      R_f[3,4] := -0.60042000;
      R_f[3,5] := 0.30684051;
      R_f[3,6] := 0.39524430;
      R_f[3,7] := 0.11368765;
      R_f[3,8] := -0.22525014;
      R_f[3,9] := 0.40331784;
      R_f[3,10] := -0.22694421;
      R_f[3,11] := 0.08383388;
      R_f[3,12] := -0.06074797;
      R_f[3,13] := -0.18165708;
      R_f[3,14] := -0.04610621;
      R_f[3,15] := -0.62458295;
      R_f[3,16] := 0.00826784;
      R_f[3,17] := 0.13735548;
      R_f[3,18] := 0.04492014;
      R_f[3,19] := -0.30372253;
      R_f[3,20] := -0.08298360;
      R_f[3,21] := 0.43319181;
      R_f[3,22] := 0.03173294;
      R_f[3,23] := 0.26679260;
      R_f[3,24] := 0.19107546;
      R_f[3,25] := -0.13225158;
      R_f[3,26] := 0.04235943;
      R_f[3,27] := 0.73829132;
      R_f[3,28] := 0.57859170;
      R_f[3,29] := -0.07161227;
      R_f[3,30] := -0.07272696;
      R_f[3,31] := -0.50867581;
      R_f[4,0] := -1.08717740;
      R_f[4,1] := -0.04287297;
      R_f[4,2] := -0.19841136;
      R_f[4,3] := 0.24848095;
      R_f[4,4] := -0.64561760;
      R_f[4,5] := -0.20718722;
      R_f[4,6] := -0.05597278;
      R_f[4,7] := -0.16602105;
      R_f[4,8] := -0.29476261;
      R_f[4,9] := 0.47976902;
      R_f[4,10] := -0.05075360;
      R_f[4,11] := 0.14082003;
      R_f[4,12] := 0.06980632;
      R_f[4,13] := 0.33018085;
      R_f[4,14] := 0.04662931;
      R_f[4,15] := -0.07799391;
      R_f[4,16] := 0.00706400;
      R_f[4,17] := 0.13971923;
      R_f[4,18] := 0.03753237;
      R_f[4,19] := -0.02597110;
      R_f[4,20] := -0.60197109;
      R_f[4,21] := 0.04454581;
      R_f[4,22] := -0.13320792;
      R_f[4,23] := 0.31133512;
      R_f[4,24] := -0.16363572;
      R_f[4,25] := 0.41873544;
      R_f[4,26] := -0.52481866;
      R_f[4,27] := 0.06860130;
      R_f[4,28] := 0.00750138;
      R_f[4,29] := 0.00922540;
      R_f[4,30] := 0.12660387;
      R_f[4,31] := 0.11132577;
      R_f[5,0] := -0.08935551;
      R_f[5,1] := 0.00341007;
      R_f[5,2] := -0.36269036;
      R_f[5,3] := -0.05915058;
      R_f[5,4] := 0.65549088;
      R_f[5,5] := -0.45446295;
      R_f[5,6] := 0.02701634;
      R_f[5,7] := 0.33505848;
      R_f[5,8] := 0.33433130;
      R_f[5,9] := -0.11102643;
      R_f[5,10] := 0.04686662;
      R_f[5,11] := -0.11728232;
      R_f[5,12] := 0.09523005;
      R_f[5,13] := -0.37170398;
      R_f[5,14] := 0.00033050;
      R_f[5,15] := 0.02845602;
      R_f[5,16] := 0.42707691;
      R_f[5,17] := -0.06965928;
      R_f[5,18] := 0.01540217;
      R_f[5,19] := -0.15121390;
      R_f[5,20] := -0.04805366;
      R_f[5,21] := -0.18535455;
      R_f[5,22] := 0.32275927;
      R_f[5,23] := -0.19729009;
      R_f[5,24] := 0.34231305;
      R_f[5,25] := -0.36576355;
      R_f[5,26] := -0.06866702;
      R_f[5,27] := 0.00050627;
      R_f[5,28] := -0.22415085;
      R_f[5,29] := 0.21506223;
      R_f[5,30] := 0.28907591;
      R_f[5,31] := 0.08619282;
      R_f[6,0] := 0.18388480;
      R_f[6,1] := 0.05767936;
      R_f[6,2] := -0.22664715;
      R_f[6,3] := 0.10472890;
      R_f[6,4] := 0.13720502;
      R_f[6,5] := -0.05844464;
      R_f[6,6] := 0.40636781;
      R_f[6,7] := 0.23722953;
      R_f[6,8] := 0.06870923;
      R_f[6,9] := -0.07299573;
      R_f[6,10] := 0.39616698;
      R_f[6,11] := 0.05431297;
      R_f[6,12] := -0.15155350;
      R_f[6,13] := -0.13813569;
      R_f[6,14] := -0.10887969;
      R_f[6,15] := -0.06144879;
      R_f[6,16] := 0.08795995;
      R_f[6,17] := -0.14627954;
      R_f[6,18] := 0.07981436;
      R_f[6,19] := 0.18627544;
      R_f[6,20] := -0.07600380;
      R_f[6,21] := -0.34014723;
      R_f[6,22] := -0.54018772;
      R_f[6,23] := 0.29552394;
      R_f[6,24] := -0.10880617;
      R_f[6,25] := -0.08422133;
      R_f[6,26] := -0.24422757;
      R_f[6,27] := -0.03805847;
      R_f[6,28] := 0.16830419;
      R_f[6,29] := -0.18664716;
      R_f[6,30] := 0.20243780;
      R_f[6,31] := 0.07874886;
      R_f[7,0] := 0.28316271;
      R_f[7,1] := 0.13009299;
      R_f[7,2] := 0.04995405;
      R_f[7,3] := 0.14345303;
      R_f[7,4] := 0.08940059;
      R_f[7,5] := -0.04840774;
      R_f[7,6] := 0.17071612;
      R_f[7,7] := -0.00365471;
      R_f[7,8] := -0.10895292;
      R_f[7,9] := -0.20513341;
      R_f[7,10] := 0.09715845;
      R_f[7,11] := 0.05839429;
      R_f[7,12] := 0.04244281;
      R_f[7,13] := -0.05333439;
      R_f[7,14] := 0.10779919;
      R_f[7,15] := 0.00831443;
      R_f[7,16] := -0.02139841;
      R_f[7,17] := -0.27714881;
      R_f[7,18] := -0.13269936;
      R_f[7,19] := 0.38708043;
      R_f[7,20] := 0.02227914;
      R_f[7,21] := -0.12789786;
      R_f[7,22] := -0.21672793;
      R_f[7,23] := 0.04945551;
      R_f[7,24] := -0.12798266;
      R_f[7,25] := -0.08468608;
      R_f[7,26] := 0.04391497;
      R_f[7,27] := 0.04113905;
      R_f[7,28] := -0.10612858;
      R_f[7,29] := 0.10980094;
      R_f[7,30] := 0.06744546;
      R_f[7,31] := 0.15760666;
      R_f[8,0] := -0.09437604;
      R_f[8,1] := 0.10058102;
      R_f[8,2] := -0.39239755;
      R_f[8,3] := 0.07142383;
      R_f[8,4] := 0.32619441;
      R_f[8,5] := -0.29801306;
      R_f[8,6] := 0.17732149;
      R_f[8,7] := 0.39382425;
      R_f[8,8] := -0.25244871;
      R_f[8,9] := -0.78001058;
      R_f[8,10] := -0.09953760;
      R_f[8,11] := -0.01873088;
      R_f[8,12] := -0.12824003;
      R_f[8,13] := -0.04000987;
      R_f[8,14] := -0.32546988;
      R_f[8,15] := -0.07414734;
      R_f[8,16] := -0.15979169;
      R_f[8,17] := -0.16899861;
      R_f[8,18] := 0.11978716;
      R_f[8,19] := -0.29437670;
      R_f[8,20] := -0.07145600;
      R_f[8,21] := 0.37895897;
      R_f[8,22] := 0.60730362;
      R_f[8,23] := -0.01808002;
      R_f[8,24] := 0.18473065;
      R_f[8,25] := -0.63517946;
      R_f[8,26] := -0.07078326;
      R_f[8,27] := 0.01834848;
      R_f[8,28] := -0.27034160;
      R_f[8,29] := 0.03424344;
      R_f[8,30] := 0.17846985;
      R_f[8,31] := -0.10791938;
      R_f[9,0] := 0.50240064;
      R_f[9,1] := -0.19293827;
      R_f[9,2] := -0.14941828;
      R_f[9,3] := 0.30088151;
      R_f[9,4] := -0.22305536;
      R_f[9,5] := -0.20884813;
      R_f[9,6] := -0.52308059;
      R_f[9,7] := -0.08416846;
      R_f[9,8] := -0.31933308;
      R_f[9,9] := 0.74035096;
      R_f[9,10] := 0.06057476;
      R_f[9,11] := -0.31038794;
      R_f[9,12] := -0.02742688;
      R_f[9,13] := 0.24148650;
      R_f[9,14] := 0.22138420;
      R_f[9,15] := -0.50248486;
      R_f[9,16] := 0.03389943;
      R_f[9,17] := -0.15244213;
      R_f[9,18] := -0.23831080;
      R_f[9,19] := 0.18266003;
      R_f[9,20] := -0.04345531;
      R_f[9,21] := -0.16341494;
      R_f[9,22] := -0.13197300;
      R_f[9,23] := -0.01865776;
      R_f[9,24] := 0.46940479;
      R_f[9,25] := 0.06735769;
      R_f[9,26] := -0.33095923;
      R_f[9,27] := -0.07481478;
      R_f[9,28] := 0.30265671;
      R_f[9,29] := -0.02983976;
      R_f[9,30] := 0.11981419;
      R_f[9,31] := 0.43036476;
      R_f[10,0] := -0.16625722;
      R_f[10,1] := 0.18885586;
      R_f[10,2] := 0.30220106;
      R_f[10,3] := -0.08386957;
      R_f[10,4] := -0.50032878;
      R_f[10,5] := 0.08482117;
      R_f[10,6] := 0.13217595;
      R_f[10,7] := 0.13670275;
      R_f[10,8] := -0.27781987;
      R_f[10,9] := 0.05184001;
      R_f[10,10] := -0.32821399;
      R_f[10,11] := 0.06394526;
      R_f[10,12] := 0.70230156;
      R_f[10,13] := 0.14407636;
      R_f[10,14] := 0.21430548;
      R_f[10,15] := -0.13537307;
      R_f[10,16] := -0.70127255;
      R_f[10,17] := 0.08713871;
      R_f[10,18] := 0.49356794;
      R_f[10,19] := -0.33338264;
      R_f[10,20] := -0.14740926;
      R_f[10,21] := 0.22738504;
      R_f[10,22] := -0.12947781;
      R_f[10,23] := 0.15810163;
      R_f[10,24] := 0.01187740;
      R_f[10,25] := 0.16353421;
      R_f[10,26] := 0.49730638;
      R_f[10,27] := -0.06625025;
      R_f[10,28] := -0.15717453;
      R_f[10,29] := -0.17355147;
      R_f[10,30] := -0.03920694;
      R_f[10,31] := 0.30297169;
      R_f[11,0] := 0.12163632;
      R_f[11,1] := -0.16561009;
      R_f[11,2] := -0.63697898;
      R_f[11,3] := -0.12967597;
      R_f[11,4] := -0.15516940;
      R_f[11,5] := -0.43934959;
      R_f[11,6] := -0.84410143;
      R_f[11,7] := -0.15710612;
      R_f[11,8] := -0.91981030;
      R_f[11,9] := 0.10710724;
      R_f[11,10] := -0.25132748;
      R_f[11,11] := 0.77600086;
      R_f[11,12] := -0.20838273;
      R_f[11,13] := 0.32214221;
      R_f[11,14] := -0.02206153;
      R_f[11,15] := -0.39864928;
      R_f[11,16] := -0.17909747;
      R_f[11,17] := -0.08701507;
      R_f[11,18] := -0.16743112;
      R_f[11,19] := -0.54472065;
      R_f[11,20] := -0.58381855;
      R_f[11,21] := 0.13781570;
      R_f[11,22] := -0.65494400;
      R_f[11,23] := 0.08265506;
      R_f[11,24] := 0.11775696;
      R_f[11,25] := 0.86460680;
      R_f[11,26] := 0.22440501;
      R_f[11,27] := 0.10443961;
      R_f[11,28] := -0.11450481;
      R_f[11,29] := 0.10720722;
      R_f[11,30] := -0.14559385;
      R_f[11,31] := -0.41325647;
      R_f[12,0] := 0.08129373;
      R_f[12,1] := 0.20157976;
      R_f[12,2] := -0.09767752;
      R_f[12,3] := 0.11404920;
      R_f[12,4] := 0.06406736;
      R_f[12,5] := -0.10172413;
      R_f[12,6] := -0.62003994;
      R_f[12,7] := 0.29222506;
      R_f[12,8] := 0.09104837;
      R_f[12,9] := 0.02718525;
      R_f[12,10] := -0.17208911;
      R_f[12,11] := 0.11898477;
      R_f[12,12] := 0.14371057;
      R_f[12,13] := 0.07740860;
      R_f[12,14] := 0.03334129;
      R_f[12,15] := -0.34480530;
      R_f[12,16] := 0.11375867;
      R_f[12,17] := -0.16553403;
      R_f[12,18] := -0.03753847;
      R_f[12,19] := 0.42828915;
      R_f[12,20] := -0.23550081;
      R_f[12,21] := -0.64313370;
      R_f[12,22] := 0.11878636;
      R_f[12,23] := 0.06645127;
      R_f[12,24] := -0.05381826;
      R_f[12,25] := -0.06362370;
      R_f[12,26] := 0.14368635;
      R_f[12,27] := 0.03581888;
      R_f[12,28] := -0.27521226;
      R_f[12,29] := -0.06815766;
      R_f[12,30] := 0.05883517;
      R_f[12,31] := 0.01413656;
      R_f[13,0] := -0.09574396;
      R_f[13,1] := 0.30759236;
      R_f[13,2] := -0.40949357;
      R_f[13,3] := -0.30002195;
      R_f[13,4] := 0.62065625;
      R_f[13,5] := -0.06791952;
      R_f[13,6] := -0.10181803;
      R_f[13,7] := 0.06609505;
      R_f[13,8] := 0.45424458;
      R_f[13,9] := -0.32844600;
      R_f[13,10] := 0.17730820;
      R_f[13,11] := -0.15458618;
      R_f[13,12] := -0.16377521;
      R_f[13,13] := 0.12967198;
      R_f[13,14] := -0.18851388;
      R_f[13,15] := 0.08791368;
      R_f[13,16] := 0.19190530;
      R_f[13,17] := -0.03352485;
      R_f[13,18] := -0.24754001;
      R_f[13,19] := -0.03332811;
      R_f[13,20] := -0.22078300;
      R_f[13,21] := -0.27547061;
      R_f[13,22] := 0.77056712;
      R_f[13,23] := -0.11708862;
      R_f[13,24] := 0.38989946;
      R_f[13,25] := 0.12295369;
      R_f[13,26] := 0.01030140;
      R_f[13,27] := -0.10658067;
      R_f[13,28] := -0.25609714;
      R_f[13,29] := 0.09743972;
      R_f[13,30] := 0.57624507;
      R_f[13,31] := 0.09921760;
      R_f[14,0] := -0.46166307;
      R_f[14,1] := -0.38297445;
      R_f[14,2] := -0.34351581;
      R_f[14,3] := 0.50245303;
      R_f[14,4] := -0.47205976;
      R_f[14,5] := -0.04034173;
      R_f[14,6] := 0.19666021;
      R_f[14,7] := -0.15099366;
      R_f[14,8] := -0.23554653;
      R_f[14,9] := 0.44932032;
      R_f[14,10] := -0.24074826;
      R_f[14,11] := 0.29974288;
      R_f[14,12] := -0.44155741;
      R_f[14,13] := 0.83714885;
      R_f[14,14] := 0.18741892;
      R_f[14,15] := -0.21850257;
      R_f[14,16] := -0.12847616;
      R_f[14,17] := 0.06488960;
      R_f[14,18] := -0.00284800;
      R_f[14,19] := -0.31293416;
      R_f[14,20] := -0.07697109;
      R_f[14,21] := 0.38044301;
      R_f[14,22] := -0.48185810;
      R_f[14,23] := -0.07073558;
      R_f[14,24] := -0.99695712;
      R_f[14,25] := 0.80939853;
      R_f[14,26] := -0.05103495;
      R_f[14,27] := -0.04504821;
      R_f[14,28] := 0.15116005;
      R_f[14,29] := -0.15104911;
      R_f[14,30] := -0.08086795;
      R_f[14,31] := -0.08960185;
      R_f[15,0] := 0.52664596;
      R_f[15,1] := 0.12164947;
      R_f[15,2] := -0.16819476;
      R_f[15,3] := -0.05969808;
      R_f[15,4] := 0.15273678;
      R_f[15,5] := -0.27137789;
      R_f[15,6] := -0.13071315;
      R_f[15,7] := 0.14372683;
      R_f[15,8] := -0.10874850;
      R_f[15,9] := 0.07457355;
      R_f[15,10] := -0.08407912;
      R_f[15,11] := 0.09970645;
      R_f[15,12] := -0.03155738;
      R_f[15,13] := -0.05560709;
      R_f[15,14] := 0.11556993;
      R_f[15,15] := -0.41232723;
      R_f[15,16] := -0.07345941;
      R_f[15,17] := 0.02771760;
      R_f[15,18] := -0.14295001;
      R_f[15,19] := -0.10515169;
      R_f[15,20] := -0.12221377;
      R_f[15,21] := -0.06810255;
      R_f[15,22] := 0.28113905;
      R_f[15,23] := -0.14406382;
      R_f[15,24] := 0.00678202;
      R_f[15,25] := -0.22208183;
      R_f[15,26] := 0.09178454;
      R_f[15,27] := -0.12816849;
      R_f[15,28] := -0.14566351;
      R_f[15,29] := -0.14765069;
      R_f[15,30] := -0.23014744;
      R_f[15,31] := -0.11258506;
      R_f[16,0] := 0.23934299;
      R_f[16,1] := -0.15829709;
      R_f[16,2] := 0.45032674;
      R_f[16,3] := 0.23261313;
      R_f[16,4] := -0.05699093;
      R_f[16,5] := -0.16829020;
      R_f[16,6] := -0.12967189;
      R_f[16,7] := 0.18884014;
      R_f[16,8] := 0.02269471;
      R_f[16,9] := 0.30370346;
      R_f[16,10] := -0.32687482;
      R_f[16,11] := 0.03308588;
      R_f[16,12] := 0.50025779;
      R_f[16,13] := 0.14397928;
      R_f[16,14] := 0.03645168;
      R_f[16,15] := -0.29107213;
      R_f[16,16] := 0.37979615;
      R_f[16,17] := 0.26871175;
      R_f[16,18] := -0.11245961;
      R_f[16,19] := -0.10605180;
      R_f[16,20] := -0.06439014;
      R_f[16,21] := -0.16872981;
      R_f[16,22] := -0.07633550;
      R_f[16,23] := -0.29030564;
      R_f[16,24] := 0.04536907;
      R_f[16,25] := -0.18899164;
      R_f[16,26] := -0.05018849;
      R_f[16,27] := -0.07462694;
      R_f[16,28] := 0.17984839;
      R_f[16,29] := -0.19122766;
      R_f[16,30] := -0.32492223;
      R_f[16,31] := -0.01023434;
      R_f[17,0] := -0.19283064;
      R_f[17,1] := 0.17507498;
      R_f[17,2] := -0.82085013;
      R_f[17,3] := 0.15822300;
      R_f[17,4] := -0.08289441;
      R_f[17,5] := -0.04341217;
      R_f[17,6] := -0.67035288;
      R_f[17,7] := -0.06796314;
      R_f[17,8] := 0.02953611;
      R_f[17,9] := 0.62533587;
      R_f[17,10] := 0.67396945;
      R_f[17,11] := 0.22164279;
      R_f[17,12] := -0.16851391;
      R_f[17,13] := 0.71597058;
      R_f[17,14] := -0.20748481;
      R_f[17,15] := 0.11059881;
      R_f[17,16] := -0.34476832;
      R_f[17,17] := 0.27433106;
      R_f[17,18] := -0.01037229;
      R_f[17,19] := -0.15571585;
      R_f[17,20] := -0.60102046;
      R_f[17,21] := 0.83061326;
      R_f[17,22] := -0.23377301;
      R_f[17,23] := -0.02111884;
      R_f[17,24] := 0.19440420;
      R_f[17,25] := 0.18241513;
      R_f[17,26] := -0.02201911;
      R_f[17,27] := -0.49202144;
      R_f[17,28] := 0.01644083;
      R_f[17,29] := -0.10121699;
      R_f[17,30] := 0.55360836;
      R_f[17,31] := -0.07391836;
      R_f[18,0] := -0.22079028;
      R_f[18,1] := -0.33156645;
      R_f[18,2] := 0.13043778;
      R_f[18,3] := 0.15372331;
      R_f[18,4] := -0.31435055;
      R_f[18,5] := -0.52705157;
      R_f[18,6] := -0.53319710;
      R_f[18,7] := -0.06062661;
      R_f[18,8] := -0.45767096;
      R_f[18,9] := 0.46125960;
      R_f[18,10] := -0.00913381;
      R_f[18,11] := 0.29711878;
      R_f[18,12] := 0.40422088;
      R_f[18,13] := 0.19489796;
      R_f[18,14] := -0.09397310;
      R_f[18,15] := 0.02433426;
      R_f[18,16] := 0.01347355;
      R_f[18,17] := 0.45005736;
      R_f[18,18] := 0.82723099;
      R_f[18,19] := 0.01506453;
      R_f[18,20] := -0.27744177;
      R_f[18,21] := 0.11534820;
      R_f[18,22] := 0.06803705;
      R_f[18,23] := -0.12547506;
      R_f[18,24] := 0.09065273;
      R_f[18,25] := -0.26198232;
      R_f[18,26] := -0.05962683;
      R_f[18,27] := -0.24309711;
      R_f[18,28] := -0.07283445;
      R_f[18,29] := 0.31726363;
      R_f[18,30] := -0.23322983;
      R_f[18,31] := -0.25323680;
      R_f[19,0] := 0.09615998;
      R_f[19,1] := 0.32398069;
      R_f[19,2] := -0.46022564;
      R_f[19,3] := 0.12604143;
      R_f[19,4] := 0.32733244;
      R_f[19,5] := -0.82866299;
      R_f[19,6] := -0.15853848;
      R_f[19,7] := -0.03126367;
      R_f[19,8] := 0.08890365;
      R_f[19,9] := -0.08684489;
      R_f[19,10] := 0.26054394;
      R_f[19,11] := -0.39950660;
      R_f[19,12] := 0.03295855;
      R_f[19,13] := -0.01441790;
      R_f[19,14] := 0.00434950;
      R_f[19,15] := -0.15201327;
      R_f[19,16] := -0.17205280;
      R_f[19,17] := -0.20647822;
      R_f[19,18] := -0.15738116;
      R_f[19,19] := -0.14136869;
      R_f[19,20] := -0.27375880;
      R_f[19,21] := -0.33055094;
      R_f[19,22] := 0.24609660;
      R_f[19,23] := -0.16637921;
      R_f[19,24] := 0.16989504;
      R_f[19,25] := 0.17177875;
      R_f[19,26] := -0.03401650;
      R_f[19,27] := -0.12747964;
      R_f[19,28] := -0.36287704;
      R_f[19,29] := -0.13957691;
      R_f[19,30] := 0.14885531;
      R_f[19,31] := 0.25682664;
      R_f[20,0] := 0.65143263;
      R_f[20,1] := 0.12967470;
      R_f[20,2] := -0.41223466;
      R_f[20,3] := -0.32649657;
      R_f[20,4] := 0.05576348;
      R_f[20,5] := -0.00373994;
      R_f[20,6] := -0.03229912;
      R_f[20,7] := 0.05183956;
      R_f[20,8] := 0.11954875;
      R_f[20,9] := -0.45034453;
      R_f[20,10] := -0.08409706;
      R_f[20,11] := -0.10399139;
      R_f[20,12] := 0.04223659;
      R_f[20,13] := -0.42114496;
      R_f[20,14] := 0.40092605;
      R_f[20,15] := 0.03704791;
      R_f[20,16] := 0.18334673;
      R_f[20,17] := -0.21014014;
      R_f[20,18] := -0.20176393;
      R_f[20,19] := 0.11477864;
      R_f[20,20] := -0.38470769;
      R_f[20,21] := -1.12075245;
      R_f[20,22] := 0.83599603;
      R_f[20,23] := 0.03310845;
      R_f[20,24] := 0.33557516;
      R_f[20,25] := -0.59122396;
      R_f[20,26] := 0.08178008;
      R_f[20,27] := -0.39574838;
      R_f[20,28] := -0.34082243;
      R_f[20,29] := 0.14776798;
      R_f[20,30] := 0.46922100;
      R_f[20,31] := 0.34887803;
      R_f[21,0] := -0.70780814;
      R_f[21,1] := -0.54152215;
      R_f[21,2] := -0.31821868;
      R_f[21,3] := 0.86289746;
      R_f[21,4] := -0.39403108;
      R_f[21,5] := -0.27079824;
      R_f[21,6] := 0.72602904;
      R_f[21,7] := 0.47715333;
      R_f[21,8] := 0.35393783;
      R_f[21,9] := -0.18864393;
      R_f[21,10] := 0.04683945;
      R_f[21,11] := -0.01854442;
      R_f[21,12] := 0.72281402;
      R_f[21,13] := 0.28782725;
      R_f[21,14] := -0.00757472;
      R_f[21,15] := -0.16304152;
      R_f[21,16] := -0.76280284;
      R_f[21,17] := 0.17034245;
      R_f[21,18] := 0.21656267;
      R_f[21,19] := -0.20434183;
      R_f[21,20] := -0.08964054;
      R_f[21,21] := 0.27781618;
      R_f[21,22] := -0.39249471;
      R_f[21,23] := 0.79524159;
      R_f[21,24] := -0.51818389;
      R_f[21,25] := 0.37090141;
      R_f[21,26] := 0.32537594;
      R_f[21,27] := -0.11953229;
      R_f[21,28] := 0.45985162;
      R_f[21,29] := 0.07980209;
      R_f[21,30] := 0.39846614;
      R_f[21,31] := -0.06241709;
      R_f[22,0] := 0.39895391;
      R_f[22,1] := 0.30520257;
      R_f[22,2] := -0.34458700;
      R_f[22,3] := -0.10527921;
      R_f[22,4] := 0.26003963;
      R_f[22,5] := -0.37983853;
      R_f[22,6] := 0.02547618;
      R_f[22,7] := -0.19680914;
      R_f[22,8] := 0.71605831;
      R_f[22,9] := 0.04098209;
      R_f[22,10] := 0.10896515;
      R_f[22,11] := -0.15730301;
      R_f[22,12] := -0.35799044;
      R_f[22,13] := -0.18627444;
      R_f[22,14] := -0.19153382;
      R_f[22,15] := -0.04852609;
      R_f[22,16] := 0.25931671;
      R_f[22,17] := -0.25600764;
      R_f[22,18] := -0.48934627;
      R_f[22,19] := -0.04790500;
      R_f[22,20] := -0.38352549;
      R_f[22,21] := -0.18561588;
      R_f[22,22] := 0.21873617;
      R_f[22,23] := 0.20801637;
      R_f[22,24] := 0.93700039;
      R_f[22,25] := 0.04714046;
      R_f[22,26] := -0.05571582;
      R_f[22,27] := 0.33375865;
      R_f[22,28] := -0.16586863;
      R_f[22,29] := -0.00929833;
      R_f[22,30] := 0.56434536;
      R_f[22,31] := 0.16850579;
      R_f[23,0] := 0.30282658;
      R_f[23,1] := -0.03574499;
      R_f[23,2] := 0.00562761;
      R_f[23,3] := 0.09418619;
      R_f[23,4] := -0.06124444;
      R_f[23,5] := -0.10330658;
      R_f[23,6] := -0.29966629;
      R_f[23,7] := 0.05105592;
      R_f[23,8] := -0.33817834;
      R_f[23,9] := -0.12041192;
      R_f[23,10] := -0.02037496;
      R_f[23,11] := 0.03016710;
      R_f[23,12] := 0.37526789;
      R_f[23,13] := 0.00504789;
      R_f[23,14] := -0.03566586;
      R_f[23,15] := -0.05691298;
      R_f[23,16] := -0.16826557;
      R_f[23,17] := 0.34201103;
      R_f[23,18] := 0.14922331;
      R_f[23,19] := 0.05192836;
      R_f[23,20] := 0.03962184;
      R_f[23,21] := -0.15185677;
      R_f[23,22] := -0.30035132;
      R_f[23,23] := 0.08715385;
      R_f[23,24] := -0.10690231;
      R_f[23,25] := -0.16740714;
      R_f[23,26] := -0.06337357;
      R_f[23,27] := -0.02622578;
      R_f[23,28] := -0.13436833;
      R_f[23,29] := 0.13256556;
      R_f[23,30] := -0.14433481;
      R_f[23,31] := 0.17851405;
      R_f[24,0] := -0.11983271;
      R_f[24,1] := 0.57634509;
      R_f[24,2] := -0.59061909;
      R_f[24,3] := -0.41855133;
      R_f[24,4] := 0.48994675;
      R_f[24,5] := -0.40760514;
      R_f[24,6] := -0.37396318;
      R_f[24,7] := 0.25456005;
      R_f[24,8] := 0.28927997;
      R_f[24,9] := -0.52789915;
      R_f[24,10] := 0.04503828;
      R_f[24,11] := -0.13581282;
      R_f[24,12] := 0.11650596;
      R_f[24,13] := -0.12701693;
      R_f[24,14] := 0.01184188;
      R_f[24,15] := -0.08589336;
      R_f[24,16] := 0.16197152;
      R_f[24,17] := -0.30688080;
      R_f[24,18] := 0.05836460;
      R_f[24,19] := -0.19957499;
      R_f[24,20] := -0.05106665;
      R_f[24,21] := -0.50352120;
      R_f[24,22] := 0.71089500;
      R_f[24,23] := -0.42265382;
      R_f[24,24] := 0.04868191;
      R_f[24,25] := -0.36235079;
      R_f[24,26] := 0.39241791;
      R_f[24,27] := -0.05973386;
      R_f[24,28] := -0.19274573;
      R_f[24,29] := 0.12360820;
      R_f[24,30] := 0.41801184;
      R_f[24,31] := -0.08968473;
      R_f[25,0] := -0.06323480;
      R_f[25,1] := 0.06630009;
      R_f[25,2] := -0.32446408;
      R_f[25,3] := 0.01768349;
      R_f[25,4] := -0.19025567;
      R_f[25,5] := -0.07292805;
      R_f[25,6] := 0.05627314;
      R_f[25,7] := -0.05622336;
      R_f[25,8] := 0.47369036;
      R_f[25,9] := -0.04888335;
      R_f[25,10] := -0.25492111;
      R_f[25,11] := -0.22475219;
      R_f[25,12] := 0.01756740;
      R_f[25,13] := 0.15392935;
      R_f[25,14] := 0.20551270;
      R_f[25,15] := -0.00423523;
      R_f[25,16] := -0.20584407;
      R_f[25,17] := -0.03102409;
      R_f[25,18] := -0.14706251;
      R_f[25,19] := 0.15027225;
      R_f[25,20] := -0.33876377;
      R_f[25,21] := -0.15575616;
      R_f[25,22] := -0.35729119;
      R_f[25,23] := -0.18495838;
      R_f[25,24] := -0.32949454;
      R_f[25,25] := 0.12997164;
      R_f[25,26] := 0.13946673;
      R_f[25,27] := -0.07950725;
      R_f[25,28] := 0.06870005;
      R_f[25,29] := 0.04001917;
      R_f[25,30] := 0.21187194;
      R_f[25,31] := -0.13515373;
      R_f[26,0] := 0.12954827;
      R_f[26,1] := 0.02364345;
      R_f[26,2] := -0.11852348;
      R_f[26,3] := -0.12563097;
      R_f[26,4] := 0.59282267;
      R_f[26,5] := -0.24795306;
      R_f[26,6] := -0.37031353;
      R_f[26,7] := 0.23576741;
      R_f[26,8] := 0.25009814;
      R_f[26,9] := -0.41952935;
      R_f[26,10] := 0.04435631;
      R_f[26,11] := -0.10239322;
      R_f[26,12] := 0.19540873;
      R_f[26,13] := -0.16128190;
      R_f[26,14] := -0.15626748;
      R_f[26,15] := -0.14187533;
      R_f[26,16] := 0.27468386;
      R_f[26,17] := 0.21832512;
      R_f[26,18] := -0.20662366;
      R_f[26,19] := -0.04332465;
      R_f[26,20] := 0.00188089;
      R_f[26,21] := -0.34826580;
      R_f[26,22] := 0.70457006;
      R_f[26,23] := -0.09021874;
      R_f[26,24] := 0.19881925;
      R_f[26,25] := -0.46599507;
      R_f[26,26] := -0.04036989;
      R_f[26,27] := 0.15067877;
      R_f[26,28] := -0.23408225;
      R_f[26,29] := -0.06713337;
      R_f[26,30] := 0.44157311;
      R_f[26,31] := 0.01604954;
      R_f[27,0] := 0.00422613;
      R_f[27,1] := -0.24214245;
      R_f[27,2] := 0.12378165;
      R_f[27,3] := 0.44537950;
      R_f[27,4] := -0.23796892;
      R_f[27,5] := -0.10803369;
      R_f[27,6] := 0.32081801;
      R_f[27,7] := 0.07398281;
      R_f[27,8] := -0.05461581;
      R_f[27,9] := 0.76077288;
      R_f[27,10] := 0.09794071;
      R_f[27,11] := 0.13426356;
      R_f[27,12] := 0.19465549;
      R_f[27,13] := 0.17829834;
      R_f[27,14] := -0.27531561;
      R_f[27,15] := 0.21807627;
      R_f[27,16] := 0.06585735;
      R_f[27,17] := 0.63826102;
      R_f[27,18] := 0.28358167;
      R_f[27,19] := 0.12067061;
      R_f[27,20] := 0.12931505;
      R_f[27,21] := 0.25539762;
      R_f[27,22] := -0.05151540;
      R_f[27,23] := 0.14127016;
      R_f[27,24] := 0.38724786;
      R_f[27,25] := -0.04042790;
      R_f[27,26] := -0.14903069;
      R_f[27,27] := 0.38932297;
      R_f[27,28] := -0.10293893;
      R_f[27,29] := 0.44895831;
      R_f[27,30] := 0.25288048;
      R_f[27,31] := -0.60808694;
      R_f[28,0] := -0.03998958;
      R_f[28,1] := 0.35614717;
      R_f[28,2] := -0.77336383;
      R_f[28,3] := -0.17002574;
      R_f[28,4] := 0.33876857;
      R_f[28,5] := -0.44312897;
      R_f[28,6] := -0.28789106;
      R_f[28,7] := -0.04398393;
      R_f[28,8] := 0.52604777;
      R_f[28,9] := 0.38523507;
      R_f[28,10] := 0.40152174;
      R_f[28,11] := -0.06791446;
      R_f[28,12] := -0.29038268;
      R_f[28,13] := 0.13817625;
      R_f[28,14] := 0.25033930;
      R_f[28,15] := -0.25225663;
      R_f[28,16] := 0.09736728;
      R_f[28,17] := -0.00644951;
      R_f[28,18] := -0.33764952;
      R_f[28,19] := -0.18797489;
      R_f[28,20] := -0.38524708;
      R_f[28,21] := -0.53872466;
      R_f[28,22] := 0.43151128;
      R_f[28,23] := -0.27624130;
      R_f[28,24] := 0.61019903;
      R_f[28,25] := 0.46353620;
      R_f[28,26] := -0.01029860;
      R_f[28,27] := -0.00695218;
      R_f[28,28] := -0.40349317;
      R_f[28,29] := 0.07006133;
      R_f[28,30] := 0.36019805;
      R_f[28,31] := 0.24174140;
      R_f[29,0] := 0.03581573;
      R_f[29,1] := -0.12398471;
      R_f[29,2] := 0.42871076;
      R_f[29,3] := -0.26184031;
      R_f[29,4] := -0.02012011;
      R_f[29,5] := -0.18130754;
      R_f[29,6] := -0.39404956;
      R_f[29,7] := 0.28413618;
      R_f[29,8] := -0.26350954;
      R_f[29,9] := 0.21336880;
      R_f[29,10] := 0.06481076;
      R_f[29,11] := 0.04123184;
      R_f[29,12] := 0.18243338;
      R_f[29,13] := -0.17203096;
      R_f[29,14] := 0.06115684;
      R_f[29,15] := -0.38312486;
      R_f[29,16] := 0.02835789;
      R_f[29,17] := 0.02435921;
      R_f[29,18] := -0.00677475;
      R_f[29,19] := -0.24558714;
      R_f[29,20] := 0.19945247;
      R_f[29,21] := 0.10431452;
      R_f[29,22] := -0.16466789;
      R_f[29,23] := 0.16764323;
      R_f[29,24] := -0.14647904;
      R_f[29,25] := -0.12140726;
      R_f[29,26] := -0.72231132;
      R_f[29,27] := -0.01095672;
      R_f[29,28] := 0.03260022;
      R_f[29,29] := -0.46683860;
      R_f[29,30] := -0.05509127;
      R_f[29,31] := -0.38489181;
      R_f[30,0] := 0.17712803;
      R_f[30,1] := -0.19013348;
      R_f[30,2] := -0.01133873;
      R_f[30,3] := 0.00156584;
      R_f[30,4] := -0.14660822;
      R_f[30,5] := -0.13482600;
      R_f[30,6] := -0.12561929;
      R_f[30,7] := 0.11202610;
      R_f[30,8] := -0.11401839;
      R_f[30,9] := 0.02297746;
      R_f[30,10] := 0.26617762;
      R_f[30,11] := 0.21258126;
      R_f[30,12] := 0.03252931;
      R_f[30,13] := -0.12060242;
      R_f[30,14] := -0.15502283;
      R_f[30,15] := -0.18934824;
      R_f[30,16] := -0.02543372;
      R_f[30,17] := 0.01465900;
      R_f[30,18] := 0.03748246;
      R_f[30,19] := -0.11580238;
      R_f[30,20] := -0.16839471;
      R_f[30,21] := -0.04181989;
      R_f[30,22] := 0.13182054;
      R_f[30,23] := -0.35960868;
      R_f[30,24] := 0.24680017;
      R_f[30,25] := -0.43622112;
      R_f[30,26] := -0.03721813;
      R_f[30,27] := -0.29478928;
      R_f[30,28] := -0.11699697;
      R_f[30,29] := 0.10289176;
      R_f[30,30] := -0.70951724;
      R_f[30,31] := 0.04023042;
      R_f[31,0] := 0.28498408;
      R_f[31,1] := -0.01036491;
      R_f[31,2] := -0.66448891;
      R_f[31,3] := 0.22786535;
      R_f[31,4] := 0.03707185;
      R_f[31,5] := -0.19638491;
      R_f[31,6] := -0.14420284;
      R_f[31,7] := 0.07611360;
      R_f[31,8] := 0.04410730;
      R_f[31,9] := -0.33191562;
      R_f[31,10] := 0.22371556;
      R_f[31,11] := -0.09215938;
      R_f[31,12] := -0.06920538;
      R_f[31,13] := -0.05639616;
      R_f[31,14] := -0.23727311;
      R_f[31,15] := -0.40676281;
      R_f[31,16] := 0.25462574;
      R_f[31,17] := -0.05670553;
      R_f[31,18] := 0.26958728;
      R_f[31,19] := 0.04933480;
      R_f[31,20] := -0.17608891;
      R_f[31,21] := 0.29653788;
      R_f[31,22] := 0.08356847;
      R_f[31,23] := -0.02820376;
      R_f[31,24] := 0.03973095;
      R_f[31,25] := -0.26713079;
      R_f[31,26] := -0.05792609;
      R_f[31,27] := -0.02376731;
      R_f[31,28] := -0.51032579;
      R_f[31,29] := -0.18555388;
      R_f[31,30] := 0.26419067;
      R_f[31,31] := -0.13750397;
      R_g[0,0] := -1.86716878;
      R_g[0,1] := 0.00594010;
      R_g[0,2] := -0.09409651;
      R_g[0,3] := -0.16056333;
      R_g[0,4] := -0.04022975;
      R_g[0,5] := -0.04449965;
      R_g[0,6] := -0.10752193;
      R_g[0,7] := -0.02334943;
      R_g[0,8] := -0.01817888;
      R_g[0,9] := -0.26527661;
      R_g[0,10] := 0.00568678;
      R_g[0,11] := 0.21044488;
      R_g[0,12] := -0.08004345;
      R_g[0,13] := 0.18242060;
      R_g[0,14] := -0.10632783;
      R_g[0,15] := 0.03126746;
      R_g[0,16] := -0.14887290;
      R_g[0,17] := 0.05704008;
      R_g[0,18] := 0.20863213;
      R_g[0,19] := -0.02117305;
      R_g[0,20] := 0.04837603;
      R_g[0,21] := -0.03557894;
      R_g[0,22] := -0.28759581;
      R_g[0,23] := 0.06040859;
      R_g[0,24] := 0.02789117;
      R_g[0,25] := 0.17847939;
      R_g[0,26] := -0.11305844;
      R_g[0,27] := -0.02103507;
      R_g[0,28] := -0.10839906;
      R_g[0,29] := -0.05569761;
      R_g[0,30] := 0.00148825;
      R_g[0,31] := 0.08525012;
      R_g[1,0] := -0.05020321;
      R_g[1,1] := -2.16353679;
      R_g[1,2] := 0.02060441;
      R_g[1,3] := -0.16821860;
      R_g[1,4] := -0.17199542;
      R_g[1,5] := -0.21708789;
      R_g[1,6] := 0.52699333;
      R_g[1,7] := 0.19596691;
      R_g[1,8] := -0.13091046;
      R_g[1,9] := -0.44146216;
      R_g[1,10] := 0.38795346;
      R_g[1,11] := 0.18625882;
      R_g[1,12] := -0.05185067;
      R_g[1,13] := 0.01474669;
      R_g[1,14] := -0.01137725;
      R_g[1,15] := -0.19595569;
      R_g[1,16] := -0.17341098;
      R_g[1,17] := 0.11021431;
      R_g[1,18] := 0.10419550;
      R_g[1,19] := -0.00315296;
      R_g[1,20] := -0.35445192;
      R_g[1,21] := 0.15130357;
      R_g[1,22] := -0.11260424;
      R_g[1,23] := -0.00286957;
      R_g[1,24] := 0.33744803;
      R_g[1,25] := 0.31054246;
      R_g[1,26] := 0.19726299;
      R_g[1,27] := -0.10143567;
      R_g[1,28] := -0.46588546;
      R_g[1,29] := 0.08564824;
      R_g[1,30] := -0.45693436;
      R_g[1,31] := 0.24614342;
      R_g[2,0] := 0.42754740;
      R_g[2,1] := -0.08439796;
      R_g[2,2] := -2.48083615;
      R_g[2,3] := 0.15594825;
      R_g[2,4] := 0.28883371;
      R_g[2,5] := -0.05249200;
      R_g[2,6] := 0.10974857;
      R_g[2,7] := 0.02201747;
      R_g[2,8] := 0.07704538;
      R_g[2,9] := -0.12673977;
      R_g[2,10] := -0.05098414;
      R_g[2,11] := -0.26468465;
      R_g[2,12] := 0.05991575;
      R_g[2,13] := -0.23358315;
      R_g[2,14] := 0.05663626;
      R_g[2,15] := -0.09780067;
      R_g[2,16] := 0.06889118;
      R_g[2,17] := 0.08715642;
      R_g[2,18] := -0.17935772;
      R_g[2,19] := 0.05660028;
      R_g[2,20] := -0.01185552;
      R_g[2,21] := 0.14994641;
      R_g[2,22] := 0.03326490;
      R_g[2,23] := -0.20292051;
      R_g[2,24] := 0.01234843;
      R_g[2,25] := -0.61469454;
      R_g[2,26] := 0.06181012;
      R_g[2,27] := 0.02427841;
      R_g[2,28] := -0.07310118;
      R_g[2,29] := -0.07686608;
      R_g[2,30] := -0.02164176;
      R_g[2,31] := -0.13903983;
      R_g[3,0] := 0.33490363;
      R_g[3,1] := -0.16903484;
      R_g[3,2] := 0.08201726;
      R_g[3,3] := 0.09150024;
      R_g[3,4] := -0.06364199;
      R_g[3,5] := 0.27780339;
      R_g[3,6] := -0.22895326;
      R_g[3,7] := 0.30511212;
      R_g[3,8] := 0.27609256;
      R_g[3,9] := -0.02962501;
      R_g[3,10] := 0.02684263;
      R_g[3,11] := 0.42021292;
      R_g[3,12] := 0.29806080;
      R_g[3,13] := 0.57169533;
      R_g[3,14] := -0.54552990;
      R_g[3,15] := -0.21052553;
      R_g[3,16] := 0.06154633;
      R_g[3,17] := 0.24341084;
      R_g[3,18] := 0.82210314;
      R_g[3,19] := 0.08356626;
      R_g[3,20] := 0.04232708;
      R_g[3,21] := -0.25469112;
      R_g[3,22] := -0.70814651;
      R_g[3,23] := 0.30768943;
      R_g[3,24] := -0.23148486;
      R_g[3,25] := 0.23140466;
      R_g[3,26] := -0.31501478;
      R_g[3,27] := 0.45398065;
      R_g[3,28] := 0.14594141;
      R_g[3,29] := -0.06619590;
      R_g[3,30] := -0.17137019;
      R_g[3,31] := 0.01482036;
      R_g[4,0] := -0.29163691;
      R_g[4,1] := 0.06742429;
      R_g[4,2] := -0.26218757;
      R_g[4,3] := -0.24882053;
      R_g[4,4] := -1.31862295;
      R_g[4,5] := 0.12687203;
      R_g[4,6] := -0.06912062;
      R_g[4,7] := -0.28659731;
      R_g[4,8] := 0.08298886;
      R_g[4,9] := 0.07161500;
      R_g[4,10] := 0.18841410;
      R_g[4,11] := 0.71728945;
      R_g[4,12] := -0.11944450;
      R_g[4,13] := -0.40399656;
      R_g[4,14] := -0.27381128;
      R_g[4,15] := 0.07633350;
      R_g[4,16] := -0.33723602;
      R_g[4,17] := 0.01599702;
      R_g[4,18] := 0.48285398;
      R_g[4,19] := -0.02277060;
      R_g[4,20] := 0.14327814;
      R_g[4,21] := -0.07385599;
      R_g[4,22] := 0.16943651;
      R_g[4,23] := 0.20791455;
      R_g[4,24] := 0.10572696;
      R_g[4,25] := -0.14309037;
      R_g[4,26] := -0.34861901;
      R_g[4,27] := -0.07557160;
      R_g[4,28] := 0.04278278;
      R_g[4,29] := 0.18120587;
      R_g[4,30] := 0.45479512;
      R_g[4,31] := 0.12026820;
      R_g[5,0] := -0.02304133;
      R_g[5,1] := 0.12000635;
      R_g[5,2] := -0.21737172;
      R_g[5,3] := 0.18598026;
      R_g[5,4] := 0.03860939;
      R_g[5,5] := -2.32899976;
      R_g[5,6] := 0.33428156;
      R_g[5,7] := 0.17339738;
      R_g[5,8] := 0.09407634;
      R_g[5,9] := -0.12730069;
      R_g[5,10] := -0.10029856;
      R_g[5,11] := 0.05282877;
      R_g[5,12] := 0.00815797;
      R_g[5,13] := 0.02642259;
      R_g[5,14] := -0.22914660;
      R_g[5,15] := 0.08215488;
      R_g[5,16] := -0.12692416;
      R_g[5,17] := 0.40874791;
      R_g[5,18] := 0.12977344;
      R_g[5,19] := -0.37322706;
      R_g[5,20] := -0.18956268;
      R_g[5,21] := 0.15636928;
      R_g[5,22] := -0.03968389;
      R_g[5,23] := 0.06268115;
      R_g[5,24] := 0.05446139;
      R_g[5,25] := 0.09671620;
      R_g[5,26] := 0.08315740;
      R_g[5,27] := 0.11672953;
      R_g[5,28] := 0.01400056;
      R_g[5,29] := -0.01500267;
      R_g[5,30] := -0.20725714;
      R_g[5,31] := -0.12881301;
      R_g[6,0] := 0.22516811;
      R_g[6,1] := 0.12028339;
      R_g[6,2] := 0.08610511;
      R_g[6,3] := 0.30619004;
      R_g[6,4] := 0.09272970;
      R_g[6,5] := -0.27587140;
      R_g[6,6] := -1.53301525;
      R_g[6,7] := 0.01461887;
      R_g[6,8] := -0.07007719;
      R_g[6,9] := -0.02174507;
      R_g[6,10] := -0.46447480;
      R_g[6,11] := -0.12738839;
      R_g[6,12] := -0.20090853;
      R_g[6,13] := 0.05110689;
      R_g[6,14] := 0.13661745;
      R_g[6,15] := -0.12478956;
      R_g[6,16] := 0.56643867;
      R_g[6,17] := -0.27863052;
      R_g[6,18] := -0.45479670;
      R_g[6,19] := -0.06489718;
      R_g[6,20] := 0.02584340;
      R_g[6,21] := -0.11935475;
      R_g[6,22] := 0.11214989;
      R_g[6,23] := -0.51340914;
      R_g[6,24] := 0.09491564;
      R_g[6,25] := -0.22439410;
      R_g[6,26] := -0.11665083;
      R_g[6,27] := -0.32614577;
      R_g[6,28] := 0.07586975;
      R_g[6,29] := -0.15533994;
      R_g[6,30] := 0.08476407;
      R_g[6,31] := 0.07970457;
      R_g[7,0] := -0.16220300;
      R_g[7,1] := 0.02679652;
      R_g[7,2] := 0.02109772;
      R_g[7,3] := -0.19320615;
      R_g[7,4] := -0.01385624;
      R_g[7,5] := -0.05546103;
      R_g[7,6] := -0.00080490;
      R_g[7,7] := -1.57574725;
      R_g[7,8] := -0.03604271;
      R_g[7,9] := 0.37345174;
      R_g[7,10] := 0.34544837;
      R_g[7,11] := 0.13587800;
      R_g[7,12] := -0.05976878;
      R_g[7,13] := -0.00776227;
      R_g[7,14] := -0.22048438;
      R_g[7,15] := 0.15726271;
      R_g[7,16] := -0.13363101;
      R_g[7,17] := 0.33995944;
      R_g[7,18] := 0.24119829;
      R_g[7,19] := 0.21298400;
      R_g[7,20] := -0.23030385;
      R_g[7,21] := -0.12107547;
      R_g[7,22] := 0.07259248;
      R_g[7,23] := 0.04259953;
      R_g[7,24] := -0.03389811;
      R_g[7,25] := 0.24742375;
      R_g[7,26] := 0.07829949;
      R_g[7,27] := 0.25065231;
      R_g[7,28] := 0.06829105;
      R_g[7,29] := 0.03315730;
      R_g[7,30] := -0.00496933;
      R_g[7,31] := -0.23368585;
      R_g[8,0] := 0.50126350;
      R_g[8,1] := -0.01075395;
      R_g[8,2] := -0.05409224;
      R_g[8,3] := -0.16767406;
      R_g[8,4] := 0.00832763;
      R_g[8,5] := 0.37799847;
      R_g[8,6] := 0.12331536;
      R_g[8,7] := -0.27819967;
      R_g[8,8] := -2.21576047;
      R_g[8,9] := 0.04844392;
      R_g[8,10] := -0.09844384;
      R_g[8,11] := 0.05162678;
      R_g[8,12] := -0.28169432;
      R_g[8,13] := -0.20529607;
      R_g[8,14] := 0.31593603;
      R_g[8,15] := 0.07457664;
      R_g[8,16] := 0.33210549;
      R_g[8,17] := -0.09959956;
      R_g[8,18] := 0.07121623;
      R_g[8,19] := 0.35284182;
      R_g[8,20] := -0.10089462;
      R_g[8,21] := -0.40786922;
      R_g[8,22] := 0.01005001;
      R_g[8,23] := 0.12587501;
      R_g[8,24] := -0.05933998;
      R_g[8,25] := 0.55777889;
      R_g[8,26] := 0.32745540;
      R_g[8,27] := 0.03045411;
      R_g[8,28] := -0.19671220;
      R_g[8,29] := -0.17951922;
      R_g[8,30] := -0.04274543;
      R_g[8,31] := 0.25599673;
      R_g[9,0] := 0.02067883;
      R_g[9,1] := 0.25770998;
      R_g[9,2] := 0.23810053;
      R_g[9,3] := 0.19122946;
      R_g[9,4] := -0.07707832;
      R_g[9,5] := 0.05503296;
      R_g[9,6] := 0.08055270;
      R_g[9,7] := 0.13022389;
      R_g[9,8] := 0.09850224;
      R_g[9,9] := -1.61873245;
      R_g[9,10] := -0.11064052;
      R_g[9,11] := 0.03935200;
      R_g[9,12] := -0.07594790;
      R_g[9,13] := 0.02672983;
      R_g[9,14] := 0.41598234;
      R_g[9,15] := -0.00220872;
      R_g[9,16] := 0.21524417;
      R_g[9,17] := -0.39857104;
      R_g[9,18] := -0.00813530;
      R_g[9,19] := -0.03940494;
      R_g[9,20] := 0.19054277;
      R_g[9,21] := 0.03413972;
      R_g[9,22] := -0.04471624;
      R_g[9,23] := -0.22795328;
      R_g[9,24] := 0.04888061;
      R_g[9,25] := -0.07975248;
      R_g[9,26] := -0.15874234;
      R_g[9,27] := -0.09421566;
      R_g[9,28] := 0.10185888;
      R_g[9,29] := -0.25601649;
      R_g[9,30] := 0.03189911;
      R_g[9,31] := 0.02803478;
      R_g[10,0] := 0.11934873;
      R_g[10,1] := -0.14988974;
      R_g[10,2] := -0.15460709;
      R_g[10,3] := -0.08242355;
      R_g[10,4] := -0.25586098;
      R_g[10,5] := -0.02314902;
      R_g[10,6] := -0.08165739;
      R_g[10,7] := 0.05377385;
      R_g[10,8] := 0.07941879;
      R_g[10,9] := -0.03854242;
      R_g[10,10] := -1.46558404;
      R_g[10,11] := 0.01830991;
      R_g[10,12] := 0.31197628;
      R_g[10,13] := -0.02278156;
      R_g[10,14] := 0.14286619;
      R_g[10,15] := -0.23215233;
      R_g[10,16] := 0.11244029;
      R_g[10,17] := -0.16206174;
      R_g[10,18] := 0.44919798;
      R_g[10,19] := 0.16908453;
      R_g[10,20] := -0.10676466;
      R_g[10,21] := 0.07486597;
      R_g[10,22] := 0.23136197;
      R_g[10,23] := 0.10003871;
      R_g[10,24] := 0.22128391;
      R_g[10,25] := -0.16353868;
      R_g[10,26] := 0.24291484;
      R_g[10,27] := 0.23580998;
      R_g[10,28] := -0.25138468;
      R_g[10,29] := 0.01641993;
      R_g[10,30] := 0.14167602;
      R_g[10,31] := 0.08870865;
      R_g[11,0] := -0.34106851;
      R_g[11,1] := -0.02875503;
      R_g[11,2] := 0.33586946;
      R_g[11,3] := 0.55462915;
      R_g[11,4] := 0.02937786;
      R_g[11,5] := 0.13981935;
      R_g[11,6] := 0.17191339;
      R_g[11,7] := -0.02137104;
      R_g[11,8] := 0.02065711;
      R_g[11,9] := -0.09035987;
      R_g[11,10] := -0.19636478;
      R_g[11,11] := -1.72786403;
      R_g[11,12] := -0.04057590;
      R_g[11,13] := 0.15109573;
      R_g[11,14] := -0.03368974;
      R_g[11,15] := -0.08068423;
      R_g[11,16] := 0.26117870;
      R_g[11,17] := 0.03805164;
      R_g[11,18] := -0.15395693;
      R_g[11,19] := -0.23101301;
      R_g[11,20] := 0.23441698;
      R_g[11,21] := -0.06810657;
      R_g[11,22] := -0.23827252;
      R_g[11,23] := -0.07978224;
      R_g[11,24] := -0.04555380;
      R_g[11,25] := -0.04114136;
      R_g[11,26] := 0.12400023;
      R_g[11,27] := 0.04892867;
      R_g[11,28] := -0.17664823;
      R_g[11,29] := -0.04479200;
      R_g[11,30] := -0.04086828;
      R_g[11,31] := 0.16403502;
      R_g[12,0] := -0.12858559;
      R_g[12,1] := 0.03379016;
      R_g[12,2] := -0.03469384;
      R_g[12,3] := 0.12741654;
      R_g[12,4] := -0.08589013;
      R_g[12,5] := -0.02192938;
      R_g[12,6] := -0.02139760;
      R_g[12,7] := -0.04024431;
      R_g[12,8] := -0.10572260;
      R_g[12,9] := -0.01926756;
      R_g[12,10] := 0.09853918;
      R_g[12,11] := 0.05490904;
      R_g[12,12] := -1.79967594;
      R_g[12,13] := -0.08506315;
      R_g[12,14] := 0.10771223;
      R_g[12,15] := 0.04973336;
      R_g[12,16] := -0.19733992;
      R_g[12,17] := 0.01932442;
      R_g[12,18] := -0.00100673;
      R_g[12,19] := -0.07807388;
      R_g[12,20] := 0.07478423;
      R_g[12,21] := 0.00233977;
      R_g[12,22] := -0.02209383;
      R_g[12,23] := 0.12203383;
      R_g[12,24] := -0.16885564;
      R_g[12,25] := 0.02344557;
      R_g[12,26] := 0.11767969;
      R_g[12,27] := 0.14465015;
      R_g[12,28] := -0.06759533;
      R_g[12,29] := 0.47032490;
      R_g[12,30] := 0.01685596;
      R_g[12,31] := -0.03329014;
      R_g[13,0] := 0.45972660;
      R_g[13,1] := 0.32463640;
      R_g[13,2] := 0.29604191;
      R_g[13,3] := 0.49243903;
      R_g[13,4] := 0.31027609;
      R_g[13,5] := -0.05934400;
      R_g[13,6] := 0.06132998;
      R_g[13,7] := 0.18528175;
      R_g[13,8] := 0.01472400;
      R_g[13,9] := -0.47797605;
      R_g[13,10] := -0.24094644;
      R_g[13,11] := -0.17913091;
      R_g[13,12] := -0.17311403;
      R_g[13,13] := -2.54636598;
      R_g[13,14] := 0.04596091;
      R_g[13,15] := -0.09920625;
      R_g[13,16] := 0.42228886;
      R_g[13,17] := 0.07932609;
      R_g[13,18] := -0.47531423;
      R_g[13,19] := -0.09417539;
      R_g[13,20] := -0.05766926;
      R_g[13,21] := -0.03843910;
      R_g[13,22] := -0.07508357;
      R_g[13,23] := -0.41806641;
      R_g[13,24] := 0.01569392;
      R_g[13,25] := 0.00260874;
      R_g[13,26] := -0.00180914;
      R_g[13,27] := -0.06168322;
      R_g[13,28] := -0.03373957;
      R_g[13,29] := -0.00371243;
      R_g[13,30] := -0.00184311;
      R_g[13,31] := 0.10216071;
      R_g[14,0] := 0.14091641;
      R_g[14,1] := 0.49853620;
      R_g[14,2] := 0.47690329;
      R_g[14,3] := 0.05769287;
      R_g[14,4] := 0.37067437;
      R_g[14,5] := 0.28377089;
      R_g[14,6] := 0.01137175;
      R_g[14,7] := -0.00710056;
      R_g[14,8] := 0.26809365;
      R_g[14,9] := -0.04161305;
      R_g[14,10] := 0.22925317;
      R_g[14,11] := -0.48795608;
      R_g[14,12] := 0.07273320;
      R_g[14,13] := 0.19280842;
      R_g[14,14] := -1.16806173;
      R_g[14,15] := -0.16170843;
      R_g[14,16] := 0.20796870;
      R_g[14,17] := 0.23254131;
      R_g[14,18] := -0.13794440;
      R_g[14,19] := -0.02917262;
      R_g[14,20] := -0.15455741;
      R_g[14,21] := -0.08204099;
      R_g[14,22] := -0.21607397;
      R_g[14,23] := -0.29174289;
      R_g[14,24] := 0.06977455;
      R_g[14,25] := -0.19362010;
      R_g[14,26] := 0.21976317;
      R_g[14,27] := 0.00026963;
      R_g[14,28] := -0.17724864;
      R_g[14,29] := 0.08898024;
      R_g[14,30] := -0.20474464;
      R_g[14,31] := 0.14378659;
      R_g[15,0] := 0.20182560;
      R_g[15,1] := 0.12131355;
      R_g[15,2] := 0.01463425;
      R_g[15,3] := 0.15993834;
      R_g[15,4] := 0.02804799;
      R_g[15,5] := -0.16840014;
      R_g[15,6] := 0.00829812;
      R_g[15,7] := 0.09067327;
      R_g[15,8] := -0.12538609;
      R_g[15,9] := -0.06829524;
      R_g[15,10] := -0.07112616;
      R_g[15,11] := -0.00371883;
      R_g[15,12] := -0.02522592;
      R_g[15,13] := -0.09582980;
      R_g[15,14] := 0.18802927;
      R_g[15,15] := -1.58931601;
      R_g[15,16] := 0.12705095;
      R_g[15,17] := -0.16617423;
      R_g[15,18] := -0.12584680;
      R_g[15,19] := -0.03204261;
      R_g[15,20] := 0.01988087;
      R_g[15,21] := 0.01436528;
      R_g[15,22] := 0.07755158;
      R_g[15,23] := 0.04729276;
      R_g[15,24] := -0.29171330;
      R_g[15,25] := -0.15872245;
      R_g[15,26] := 0.18300183;
      R_g[15,27] := -0.08073322;
      R_g[15,28] := -0.04181913;
      R_g[15,29] := -0.23932807;
      R_g[15,30] := -0.07486971;
      R_g[15,31] := 0.10602318;
      R_g[16,0] := -0.06681629;
      R_g[16,1] := 0.07036684;
      R_g[16,2] := -0.05912037;
      R_g[16,3] := 0.08132802;
      R_g[16,4] := 0.11257288;
      R_g[16,5] := 0.09455875;
      R_g[16,6] := -0.34879151;
      R_g[16,7] := -0.04252379;
      R_g[16,8] := -0.03194689;
      R_g[16,9] := 0.00343745;
      R_g[16,10] := -0.15653400;
      R_g[16,11] := -0.14295644;
      R_g[16,12] := -0.02853871;
      R_g[16,13] := -0.10090829;
      R_g[16,14] := 0.03872371;
      R_g[16,15] := 0.24959658;
      R_g[16,16] := -1.38679147;
      R_g[16,17] := -0.03435654;
      R_g[16,18] := -0.15214655;
      R_g[16,19] := 0.00448510;
      R_g[16,20] := 0.10372234;
      R_g[16,21] := 0.29237437;
      R_g[16,22] := -0.00143967;
      R_g[16,23] := 0.05745683;
      R_g[16,24] := -0.13639535;
      R_g[16,25] := 0.15248059;
      R_g[16,26] := 0.07691783;
      R_g[16,27] := -0.13439301;
      R_g[16,28] := -0.08911712;
      R_g[16,29] := -0.06526610;
      R_g[16,30] := 0.33859855;
      R_g[16,31] := 0.14029105;
      R_g[17,0] := 0.14671518;
      R_g[17,1] := -0.20630203;
      R_g[17,2] := 0.68066353;
      R_g[17,3] := 0.41419700;
      R_g[17,4] := -0.16559522;
      R_g[17,5] := 0.03802754;
      R_g[17,6] := -0.10850023;
      R_g[17,7] := -0.10096590;
      R_g[17,8] := -0.47244051;
      R_g[17,9] := 0.45527029;
      R_g[17,10] := -0.35605320;
      R_g[17,11] := 0.05101961;
      R_g[17,12] := -0.39417115;
      R_g[17,13] := 0.39322102;
      R_g[17,14] := -0.09366875;
      R_g[17,15] := -0.30847651;
      R_g[17,16] := 0.40280735;
      R_g[17,17] := -1.18712938;
      R_g[17,18] := -0.24961938;
      R_g[17,19] := -0.39374694;
      R_g[17,20] := -0.00170897;
      R_g[17,21] := 0.39039624;
      R_g[17,22] := -0.92846608;
      R_g[17,23] := -0.07637399;
      R_g[17,24] := -0.32924676;
      R_g[17,25] := 0.03110591;
      R_g[17,26] := 0.04365248;
      R_g[17,27] := 0.14979164;
      R_g[17,28] := 0.07266354;
      R_g[17,29] := -0.01802464;
      R_g[17,30] := -0.12855233;
      R_g[17,31] := -0.13632473;
      R_g[18,0] := 0.61803639;
      R_g[18,1] := 0.25511530;
      R_g[18,2] := 0.05195731;
      R_g[18,3] := 0.37520856;
      R_g[18,4] := 0.39242169;
      R_g[18,5] := -0.10294182;
      R_g[18,6] := 0.26254231;
      R_g[18,7] := 0.04468368;
      R_g[18,8] := -0.03643387;
      R_g[18,9] := -0.31122327;
      R_g[18,10] := -0.00521892;
      R_g[18,11] := -0.20397757;
      R_g[18,12] := -0.24374188;
      R_g[18,13] := 0.22966601;
      R_g[18,14] := -0.00486043;
      R_g[18,15] := -0.29596737;
      R_g[18,16] := 0.26810029;
      R_g[18,17] := 0.19241925;
      R_g[18,18] := -1.71501064;
      R_g[18,19] := 0.04475369;
      R_g[18,20] := -0.14080441;
      R_g[18,21] := 0.19410335;
      R_g[18,22] := 0.04632924;
      R_g[18,23] := -0.19822948;
      R_g[18,24] := -0.01822053;
      R_g[18,25] := 0.00715217;
      R_g[18,26] := 0.05302840;
      R_g[18,27] := 0.04905124;
      R_g[18,28] := -0.07875889;
      R_g[18,29] := -0.02230844;
      R_g[18,30] := 0.04014237;
      R_g[18,31] := -0.02884550;
      R_g[19,0] := -0.75135368;
      R_g[19,1] := -0.21284764;
      R_g[19,2] := -0.19804505;
      R_g[19,3] := -0.12862568;
      R_g[19,4] := -0.46584809;
      R_g[19,5] := -0.05286160;
      R_g[19,6] := -0.10783059;
      R_g[19,7] := 0.04422674;
      R_g[19,8] := 0.03374076;
      R_g[19,9] := 0.01016540;
      R_g[19,10] := -0.18281689;
      R_g[19,11] := 0.27606329;
      R_g[19,12] := -0.06603118;
      R_g[19,13] := -0.01851949;
      R_g[19,14] := -0.35077471;
      R_g[19,15] := 0.24131002;
      R_g[19,16] := -0.37709793;
      R_g[19,17] := 0.35459128;
      R_g[19,18] := 0.37763101;
      R_g[19,19] := -2.10741782;
      R_g[19,20] := -0.13689831;
      R_g[19,21] := 0.01539214;
      R_g[19,22] := -0.00843668;
      R_g[19,23] := 0.53741390;
      R_g[19,24] := -0.10536232;
      R_g[19,25] := 0.10730530;
      R_g[19,26] := -0.13406259;
      R_g[19,27] := 0.27381045;
      R_g[19,28] := 0.00509977;
      R_g[19,29] := 0.18445835;
      R_g[19,30] := -0.01738629;
      R_g[19,31] := -0.06444063;
      R_g[20,0] := 0.18924890;
      R_g[20,1] := 0.18402432;
      R_g[20,2] := 0.02781527;
      R_g[20,3] := 0.23947574;
      R_g[20,4] := -0.08406357;
      R_g[20,5] := 0.12817335;
      R_g[20,6] := 0.30762580;
      R_g[20,7] := 0.04187437;
      R_g[20,8] := 0.27227950;
      R_g[20,9] := -0.11457944;
      R_g[20,10] := -0.20207560;
      R_g[20,11] := 0.09050925;
      R_g[20,12] := -0.10230012;
      R_g[20,13] := 0.18245421;
      R_g[20,14] := 0.14094315;
      R_g[20,15] := -0.21245943;
      R_g[20,16] := 0.22506553;
      R_g[20,17] := -0.03114314;
      R_g[20,18] := 0.25464541;
      R_g[20,19] := 0.15946212;
      R_g[20,20] := -2.75024509;
      R_g[20,21] := 0.01992022;
      R_g[20,22] := 0.03351297;
      R_g[20,23] := -0.30453184;
      R_g[20,24] := 0.15048067;
      R_g[20,25] := 0.03220677;
      R_g[20,26] := 0.14691569;
      R_g[20,27] := 0.20233470;
      R_g[20,28] := -0.11183912;
      R_g[20,29] := 0.00709963;
      R_g[20,30] := -0.10263816;
      R_g[20,31] := -0.11027271;
      R_g[21,0] := -0.08157737;
      R_g[21,1] := 0.12452888;
      R_g[21,2] := -0.07601022;
      R_g[21,3] := 0.25199667;
      R_g[21,4] := 0.06423903;
      R_g[21,5] := 0.12198128;
      R_g[21,6] := -0.47932604;
      R_g[21,7] := -0.05985606;
      R_g[21,8] := 0.22486039;
      R_g[21,9] := -0.00334445;
      R_g[21,10] := -0.23857601;
      R_g[21,11] := -0.02146066;
      R_g[21,12] := -0.28514680;
      R_g[21,13] := 0.11122446;
      R_g[21,14] := -0.24231751;
      R_g[21,15] := -0.17232344;
      R_g[21,16] := 0.30115235;
      R_g[21,17] := 0.11670188;
      R_g[21,18] := -0.03272144;
      R_g[21,19] := -0.14810626;
      R_g[21,20] := 0.14458667;
      R_g[21,21] := -0.53038293;
      R_g[21,22] := -0.18996024;
      R_g[21,23] := -0.07745564;
      R_g[21,24] := 0.21534516;
      R_g[21,25] := -0.13944361;
      R_g[21,26] := -0.20756353;
      R_g[21,27] := 0.23508912;
      R_g[21,28] := -0.00923094;
      R_g[21,29] := 0.03929158;
      R_g[21,30] := 0.07484641;
      R_g[21,31] := -0.02914809;
      R_g[22,0] := 0.50535607;
      R_g[22,1] := -0.06260853;
      R_g[22,2] := 0.08109864;
      R_g[22,3] := 0.01245827;
      R_g[22,4] := 0.23083940;
      R_g[22,5] := -0.09113465;
      R_g[22,6] := 0.01330733;
      R_g[22,7] := 0.10156141;
      R_g[22,8] := -0.09307987;
      R_g[22,9] := -0.20655596;
      R_g[22,10] := -0.51928091;
      R_g[22,11] := -0.15207466;
      R_g[22,12] := -0.06335686;
      R_g[22,13] := 0.07315928;
      R_g[22,14] := 0.32269958;
      R_g[22,15] := -0.09189125;
      R_g[22,16] := 0.40304139;
      R_g[22,17] := -0.40450314;
      R_g[22,18] := -0.63684171;
      R_g[22,19] := -0.15540077;
      R_g[22,20] := 0.00914839;
      R_g[22,21] := 0.08185407;
      R_g[22,22] := -2.49282122;
      R_g[22,23] := -0.38054550;
      R_g[22,24] := -0.00924153;
      R_g[22,25] := -0.00120828;
      R_g[22,26] := -0.20842904;
      R_g[22,27] := -0.15960918;
      R_g[22,28] := -0.16979735;
      R_g[22,29] := 0.04954208;
      R_g[22,30] := 0.10421277;
      R_g[22,31] := 0.10225163;
      R_g[23,0] := 0.18052800;
      R_g[23,1] := -0.07720698;
      R_g[23,2] := 0.15911111;
      R_g[23,3] := 0.30997247;
      R_g[23,4] := 0.16866267;
      R_g[23,5] := 0.00785692;
      R_g[23,6] := 0.00494674;
      R_g[23,7] := -0.06666262;
      R_g[23,8] := 0.06490348;
      R_g[23,9] := -0.19479643;
      R_g[23,10] := -0.14945234;
      R_g[23,11] := -0.05691649;
      R_g[23,12] := -0.21839225;
      R_g[23,13] := 0.22376211;
      R_g[23,14] := 0.01327592;
      R_g[23,15] := 0.19760872;
      R_g[23,16] := 0.07945457;
      R_g[23,17] := -0.01825088;
      R_g[23,18] := -0.14043757;
      R_g[23,19] := 0.00620574;
      R_g[23,20] := 0.09369237;
      R_g[23,21] := -0.03980252;
      R_g[23,22] := 0.19607799;
      R_g[23,23] := -1.43363607;
      R_g[23,24] := 0.02975971;
      R_g[23,25] := -0.16353932;
      R_g[23,26] := -0.12808764;
      R_g[23,27] := -0.14395322;
      R_g[23,28] := -0.09217037;
      R_g[23,29] := 0.24549456;
      R_g[23,30] := 0.10042652;
      R_g[23,31] := 0.08094314;
      R_g[24,0] := -0.26641947;
      R_g[24,1] := -0.23788896;
      R_g[24,2] := 0.26894578;
      R_g[24,3] := -0.32378414;
      R_g[24,4] := -0.04978346;
      R_g[24,5] := 0.09013753;
      R_g[24,6] := -0.10760899;
      R_g[24,7] := 0.04824702;
      R_g[24,8] := -0.10581810;
      R_g[24,9] := 0.15669861;
      R_g[24,10] := 0.12566140;
      R_g[24,11] := -0.04599889;
      R_g[24,12] := 0.24090631;
      R_g[24,13] := 0.03215941;
      R_g[24,14] := 0.05187291;
      R_g[24,15] := 0.26031712;
      R_g[24,16] := -0.21561927;
      R_g[24,17] := -0.02364190;
      R_g[24,18] := 0.09312176;
      R_g[24,19] := 0.13471472;
      R_g[24,20] := 0.29225814;
      R_g[24,21] := 0.04183585;
      R_g[24,22] := -0.06511365;
      R_g[24,23] := 0.14407112;
      R_g[24,24] := -2.98465896;
      R_g[24,25] := -0.10412049;
      R_g[24,26] := -0.19039965;
      R_g[24,27] := -0.04051330;
      R_g[24,28] := 0.00060194;
      R_g[24,29] := 0.16535380;
      R_g[24,30] := 0.04648554;
      R_g[24,31] := -0.02625122;
      R_g[25,0] := 0.43024307;
      R_g[25,1] := 0.10947325;
      R_g[25,2] := -0.03608720;
      R_g[25,3] := 0.22247598;
      R_g[25,4] := 0.44687057;
      R_g[25,5] := 0.02062996;
      R_g[25,6] := 0.03161010;
      R_g[25,7] := -0.05541447;
      R_g[25,8] := -0.08682021;
      R_g[25,9] := -0.20357162;
      R_g[25,10] := 0.16417988;
      R_g[25,11] := -0.26040092;
      R_g[25,12] := -0.14754145;
      R_g[25,13] := 0.13008007;
      R_g[25,14] := -0.29289693;
      R_g[25,15] := -0.15000887;
      R_g[25,16] := 0.17711322;
      R_g[25,17] := 0.04820256;
      R_g[25,18] := -0.30309179;
      R_g[25,19] := -0.09854405;
      R_g[25,20] := 0.08423353;
      R_g[25,21] := -0.07758698;
      R_g[25,22] := 0.00059808;
      R_g[25,23] := -0.14276446;
      R_g[25,24] := -0.09778740;
      R_g[25,25] := -1.41535318;
      R_g[25,26] := 0.07131358;
      R_g[25,27] := 0.04293850;
      R_g[25,28] := 0.12346980;
      R_g[25,29] := -0.06572708;
      R_g[25,30] := -0.04491949;
      R_g[25,31] := 0.06688137;
      R_g[26,0] := 0.24152957;
      R_g[26,1] := 0.01735749;
      R_g[26,2] := 0.04355362;
      R_g[26,3] := 0.06117517;
      R_g[26,4] := 0.32630402;
      R_g[26,5] := 0.07351752;
      R_g[26,6] := 0.06187835;
      R_g[26,7] := -0.09732439;
      R_g[26,8] := 0.28992870;
      R_g[26,9] := 0.16822580;
      R_g[26,10] := 0.16118686;
      R_g[26,11] := -0.10133380;
      R_g[26,12] := -0.04566494;
      R_g[26,13] := -0.03849275;
      R_g[26,14] := -0.06276733;
      R_g[26,15] := 0.00862427;
      R_g[26,16] := 0.06850542;
      R_g[26,17] := 0.06419130;
      R_g[26,18] := 0.03335274;
      R_g[26,19] := 0.19523142;
      R_g[26,20] := 0.49831131;
      R_g[26,21] := 0.01160550;
      R_g[26,22] := 0.03584570;
      R_g[26,23] := -0.09505314;
      R_g[26,24] := -0.19243982;
      R_g[26,25] := -0.47533280;
      R_g[26,26] := -2.50729489;
      R_g[26,27] := 0.00985446;
      R_g[26,28] := 0.01180097;
      R_g[26,29] := -0.28736252;
      R_g[26,30] := -0.02167805;
      R_g[26,31] := -0.11752307;
      R_g[27,0] := 0.01092918;
      R_g[27,1] := 0.18430310;
      R_g[27,2] := 0.06490619;
      R_g[27,3] := 0.29795435;
      R_g[27,4] := 0.01091339;
      R_g[27,5] := -0.02555788;
      R_g[27,6] := 0.04701962;
      R_g[27,7] := 0.25866464;
      R_g[27,8] := -0.05091048;
      R_g[27,9] := -0.12615849;
      R_g[27,10] := 0.22210193;
      R_g[27,11] := -0.02660196;
      R_g[27,12] := 0.35353318;
      R_g[27,13] := -0.05878561;
      R_g[27,14] := 0.02708012;
      R_g[27,15] := -0.34227443;
      R_g[27,16] := 0.16814435;
      R_g[27,17] := -0.06724432;
      R_g[27,18] := -0.23303925;
      R_g[27,19] := -0.19293629;
      R_g[27,20] := -0.09463950;
      R_g[27,21] := 0.08244657;
      R_g[27,22] := -0.27527824;
      R_g[27,23] := -0.05257547;
      R_g[27,24] := -0.00907461;
      R_g[27,25] := 0.11327704;
      R_g[27,26] := 0.17048852;
      R_g[27,27] := -1.01607871;
      R_g[27,28] := 0.24251650;
      R_g[27,29] := -0.47379026;
      R_g[27,30] := -0.06415563;
      R_g[27,31] := 0.21514556;
      R_g[28,0] := 0.20224625;
      R_g[28,1] := 0.19573490;
      R_g[28,2] := 0.01332051;
      R_g[28,3] := 0.46680877;
      R_g[28,4] := 0.23773916;
      R_g[28,5] := 0.32944795;
      R_g[28,6] := -0.24991669;
      R_g[28,7] := 0.10101810;
      R_g[28,8] := 0.14906435;
      R_g[28,9] := -0.07248143;
      R_g[28,10] := -0.22717230;
      R_g[28,11] := -0.16842264;
      R_g[28,12] := -0.43922180;
      R_g[28,13] := -0.01462650;
      R_g[28,14] := 0.01292261;
      R_g[28,15] := 0.07795207;
      R_g[28,16] := 0.29460794;
      R_g[28,17] := 0.41332749;
      R_g[28,18] := -0.21009579;
      R_g[28,19] := 0.42963541;
      R_g[28,20] := 0.00025508;
      R_g[28,21] := -0.10620708;
      R_g[28,22] := 0.17958641;
      R_g[28,23] := 0.02184093;
      R_g[28,24] := -0.40841687;
      R_g[28,25] := -0.25509256;
      R_g[28,26] := -0.17728026;
      R_g[28,27] := 0.11402236;
      R_g[28,28] := -3.10649037;
      R_g[28,29] := -0.36601931;
      R_g[28,30] := 0.08261382;
      R_g[28,31] := -0.49876866;
      R_g[29,0] := -0.18599495;
      R_g[29,1] := -0.30418199;
      R_g[29,2] := 0.11100125;
      R_g[29,3] := -0.05784649;
      R_g[29,4] := 0.10008840;
      R_g[29,5] := 0.08896575;
      R_g[29,6] := 0.30683702;
      R_g[29,7] := -0.16360219;
      R_g[29,8] := 0.13722138;
      R_g[29,9] := 0.15708315;
      R_g[29,10] := 0.33288050;
      R_g[29,11] := 0.02937395;
      R_g[29,12] := 0.04896364;
      R_g[29,13] := 0.00104734;
      R_g[29,14] := -0.16367893;
      R_g[29,15] := 0.16312605;
      R_g[29,16] := -0.13079922;
      R_g[29,17] := 0.26347440;
      R_g[29,18] := -0.09648097;
      R_g[29,19] := 0.31666356;
      R_g[29,20] := -0.28754526;
      R_g[29,21] := 0.18227148;
      R_g[29,22] := 0.15559122;
      R_g[29,23] := -0.14756282;
      R_g[29,24] := -0.01094520;
      R_g[29,25] := 0.01550437;
      R_g[29,26] := 0.27994382;
      R_g[29,27] := 0.07359030;
      R_g[29,28] := 0.00251217;
      R_g[29,29] := -1.41211045;
      R_g[29,30] := -0.04146304;
      R_g[29,31] := -0.34272864;
      R_g[30,0] := -0.05406943;
      R_g[30,1] := 0.11439317;
      R_g[30,2] := -0.16407579;
      R_g[30,3] := -0.06813712;
      R_g[30,4] := -0.03963117;
      R_g[30,5] := -0.09176665;
      R_g[30,6] := 0.05011456;
      R_g[30,7] := 0.01465930;
      R_g[30,8] := -0.19538324;
      R_g[30,9] := 0.00951732;
      R_g[30,10] := 0.25830692;
      R_g[30,11] := -0.12469292;
      R_g[30,12] := 0.08887242;
      R_g[30,13] := -0.12981550;
      R_g[30,14] := 0.14200117;
      R_g[30,15] := -0.16436660;
      R_g[30,16] := -0.33510593;
      R_g[30,17] := 0.02839339;
      R_g[30,18] := 0.18479024;
      R_g[30,19] := -0.06274416;
      R_g[30,20] := -0.06184945;
      R_g[30,21] := 0.04965051;
      R_g[30,22] := 0.00922537;
      R_g[30,23] := 0.01295749;
      R_g[30,24] := 0.10369122;
      R_g[30,25] := 0.14547619;
      R_g[30,26] := 0.09004135;
      R_g[30,27] := -0.06731008;
      R_g[30,28] := 0.01577213;
      R_g[30,29] := 0.00694244;
      R_g[30,30] := -1.30016100;
      R_g[30,31] := 0.04289828;
      R_g[31,0] := 0.25758705;
      R_g[31,1] := 0.03670706;
      R_g[31,2] := -0.32024196;
      R_g[31,3] := 0.44765759;
      R_g[31,4] := 0.21751612;
      R_g[31,5] := 0.23459953;
      R_g[31,6] := -0.12392062;
      R_g[31,7] := 0.04603523;
      R_g[31,8] := 0.16177517;
      R_g[31,9] := -0.48068467;
      R_g[31,10] := -0.20070654;
      R_g[31,11] := -0.14613695;
      R_g[31,12] := -0.54277533;
      R_g[31,13] := -0.07106268;
      R_g[31,14] := -0.41382626;
      R_g[31,15] := 0.20374061;
      R_g[31,16] := 0.05723839;
      R_g[31,17] := -0.04078045;
      R_g[31,18] := 0.16072863;
      R_g[31,19] := -0.03207170;
      R_g[31,20] := 0.01617512;
      R_g[31,21] := -0.08424362;
      R_g[31,22] := 0.14073916;
      R_g[31,23] := -0.06544417;
      R_g[31,24] := 0.34330231;
      R_g[31,25] := -0.19045305;
      R_g[31,26] := 0.30024353;
      R_g[31,27] := 0.06452943;
      R_g[31,28] := 0.26819456;
      R_g[31,29] := -0.23753491;
      R_g[31,30] := 0.12559205;
      R_g[31,31] := -1.87869716;
      R_o[0,0] := 1.04179561;
      R_o[0,1] := 0.92017525;
      R_o[0,2] := -1.79505873;
      R_o[0,3] := -0.19103914;
      R_o[0,4] := 0.95653963;
      R_o[0,5] := -0.53679043;
      R_o[0,6] := 0.13910255;
      R_o[0,7] := 0.36717987;
      R_o[0,8] := 0.13132155;
      R_o[0,9] := -0.51269883;
      R_o[0,10] := -0.05477599;
      R_o[0,11] := -0.67714477;
      R_o[0,12] := -0.07006622;
      R_o[0,13] := -1.38233066;
      R_o[0,14] := 0.61216694;
      R_o[0,15] := -0.03455535;
      R_o[0,16] := 0.39541319;
      R_o[0,17] := -0.81024104;
      R_o[0,18] := -0.38071778;
      R_o[0,19] := 0.33111337;
      R_o[0,20] := -0.56832236;
      R_o[0,21] := -0.18811585;
      R_o[0,22] := 0.99759519;
      R_o[0,23] := -0.46505177;
      R_o[0,24] := 1.28675437;
      R_o[0,25] := -0.28324643;
      R_o[0,26] := 0.11801465;
      R_o[0,27] := -0.49335349;
      R_o[0,28] := -0.16024339;
      R_o[0,29] := 0.00303155;
      R_o[0,30] := -0.07324440;
      R_o[0,31] := 1.07838094;
      R_o[1,0] := -0.17481463;
      R_o[1,1] := -0.90838975;
      R_o[1,2] := -0.54029238;
      R_o[1,3] := -0.30299738;
      R_o[1,4] := 0.37807101;
      R_o[1,5] := -0.37692639;
      R_o[1,6] := -0.21153799;
      R_o[1,7] := -0.23047979;
      R_o[1,8] := 0.43772149;
      R_o[1,9] := -0.13093925;
      R_o[1,10] := 0.00866629;
      R_o[1,11] := -0.03386870;
      R_o[1,12] := 0.35904413;
      R_o[1,13] := -0.54963106;
      R_o[1,14] := -0.15785606;
      R_o[1,15] := 0.64084804;
      R_o[1,16] := 0.01572920;
      R_o[1,17] := -0.48720333;
      R_o[1,18] := -0.17887083;
      R_o[1,19] := 0.31963482;
      R_o[1,20] := -0.28216973;
      R_o[1,21] := -0.59497058;
      R_o[1,22] := 0.60120654;
      R_o[1,23] := -0.27428257;
      R_o[1,24] := 0.50388652;
      R_o[1,25] := 0.16748510;
      R_o[1,26] := -0.04107720;
      R_o[1,27] := -0.57918507;
      R_o[1,28] := 0.20662229;
      R_o[1,29] := 0.14393075;
      R_o[1,30] := -0.01422888;
      R_o[1,31] := 0.09393608;
      R_o[2,0] := -0.06871614;
      R_o[2,1] := 0.63711506;
      R_o[2,2] := -0.38377136;
      R_o[2,3] := -0.17974423;
      R_o[2,4] := 0.32400796;
      R_o[2,5] := -0.03171432;
      R_o[2,6] := -0.29403153;
      R_o[2,7] := 0.06398765;
      R_o[2,8] := 0.17373838;
      R_o[2,9] := -0.15972729;
      R_o[2,10] := 0.45576304;
      R_o[2,11] := -0.93120134;
      R_o[2,12] := 0.04551729;
      R_o[2,13] := -0.87977225;
      R_o[2,14] := -0.25093880;
      R_o[2,15] := 0.39677525;
      R_o[2,16] := 0.01663817;
      R_o[2,17] := -0.77001494;
      R_o[2,18] := -0.18905999;
      R_o[2,19] := 0.04578963;
      R_o[2,20] := -0.00495861;
      R_o[2,21] := -0.14044468;
      R_o[2,22] := 0.27766317;
      R_o[2,23] := -0.37402457;
      R_o[2,24] := 1.21451783;
      R_o[2,25] := -0.42607296;
      R_o[2,26] := 0.33055431;
      R_o[2,27] := -0.68634737;
      R_o[2,28] := -0.52980918;
      R_o[2,29] := 0.61272937;
      R_o[2,30] := 0.24327858;
      R_o[2,31] := 0.19622318;
      R_o[3,0] := -0.17584245;
      R_o[3,1] := -0.17390651;
      R_o[3,2] := -0.00588614;
      R_o[3,3] := 0.78035086;
      R_o[3,4] := -0.32025203;
      R_o[3,5] := 0.23440066;
      R_o[3,6] := 0.49464506;
      R_o[3,7] := 0.04548555;
      R_o[3,8] := 0.05832842;
      R_o[3,9] := 0.00163286;
      R_o[3,10] := 0.15238303;
      R_o[3,11] := -0.23099470;
      R_o[3,12] := -0.08316677;
      R_o[3,13] := -0.29882267;
      R_o[3,14] := 0.28996965;
      R_o[3,15] := 0.01960599;
      R_o[3,16] := 0.15619060;
      R_o[3,17] := 0.24800168;
      R_o[3,18] := -0.31017816;
      R_o[3,19] := 0.14146750;
      R_o[3,20] := -0.03939479;
      R_o[3,21] := 0.15289256;
      R_o[3,22] := 0.40393239;
      R_o[3,23] := 0.00665908;
      R_o[3,24] := -0.04982851;
      R_o[3,25] := -0.41707465;
      R_o[3,26] := 0.20472930;
      R_o[3,27] := -0.14279339;
      R_o[3,28] := -0.04745095;
      R_o[3,29] := 0.23318978;
      R_o[3,30] := 0.24752939;
      R_o[3,31] := -0.02279269;
      R_o[4,0] := 0.28966746;
      R_o[4,1] := 0.24345395;
      R_o[4,2] := -0.23835556;
      R_o[4,3] := -0.18675509;
      R_o[4,4] := -1.14337611;
      R_o[4,5] := 0.03564367;
      R_o[4,6] := 0.25256306;
      R_o[4,7] := -0.18545251;
      R_o[4,8] := 0.21089309;
      R_o[4,9] := -0.51671422;
      R_o[4,10] := -0.27655339;
      R_o[4,11] := -0.21483746;
      R_o[4,12] := -0.24700516;
      R_o[4,13] := -0.23963267;
      R_o[4,14] := -0.93672627;
      R_o[4,15] := 0.06121854;
      R_o[4,16] := -0.03358792;
      R_o[4,17] := -0.09474288;
      R_o[4,18] := -0.03891778;
      R_o[4,19] := 0.14612053;
      R_o[4,20] := -0.09566169;
      R_o[4,21] := -0.05828689;
      R_o[4,22] := 0.15136474;
      R_o[4,23] := -0.19155599;
      R_o[4,24] := 0.14552544;
      R_o[4,25] := 0.57355893;
      R_o[4,26] := 0.03241645;
      R_o[4,27] := -0.26198941;
      R_o[4,28] := 0.20363624;
      R_o[4,29] := 0.38784343;
      R_o[4,30] := 0.13299167;
      R_o[4,31] := 0.05830654;
      R_o[5,0] := 0.28887334;
      R_o[5,1] := 0.20251507;
      R_o[5,2] := -0.81091332;
      R_o[5,3] := -0.63600522;
      R_o[5,4] := 0.67597026;
      R_o[5,5] := -0.39085054;
      R_o[5,6] := -0.23710330;
      R_o[5,7] := -0.01203742;
      R_o[5,8] := 1.16759574;
      R_o[5,9] := -0.52899224;
      R_o[5,10] := 0.19900157;
      R_o[5,11] := -0.63206440;
      R_o[5,12] := 0.04855163;
      R_o[5,13] := -0.89585042;
      R_o[5,14] := 0.05872724;
      R_o[5,15] := 0.84902614;
      R_o[5,16] := -0.01854324;
      R_o[5,17] := -0.50847763;
      R_o[5,18] := -0.13442311;
      R_o[5,19] := -0.09384207;
      R_o[5,20] := -0.22825406;
      R_o[5,21] := -1.27563584;
      R_o[5,22] := 0.47145090;
      R_o[5,23] := -0.05726700;
      R_o[5,24] := 1.12635720;
      R_o[5,25] := -0.30669662;
      R_o[5,26] := 0.31779301;
      R_o[5,27] := 0.10437986;
      R_o[5,28] := -0.36161882;
      R_o[5,29] := 0.34370479;
      R_o[5,30] := 0.32471529;
      R_o[5,31] := 0.62782931;
      R_o[6,0] := -0.02902499;
      R_o[6,1] := 0.31040263;
      R_o[6,2] := -0.03964311;
      R_o[6,3] := -0.17946681;
      R_o[6,4] := 0.25533327;
      R_o[6,5] := 0.36727500;
      R_o[6,6] := -0.32601824;
      R_o[6,7] := -0.23880924;
      R_o[6,8] := 0.27495176;
      R_o[6,9] := -0.08483669;
      R_o[6,10] := 0.25587347;
      R_o[6,11] := -0.13982451;
      R_o[6,12] := -0.10905550;
      R_o[6,13] := -0.41834557;
      R_o[6,14] := -0.59158003;
      R_o[6,15] := 0.26055050;
      R_o[6,16] := 0.19347337;
      R_o[6,17] := -0.18370837;
      R_o[6,18] := -0.03631273;
      R_o[6,19] := 0.00060258;
      R_o[6,20] := -0.13735239;
      R_o[6,21] := 0.01526413;
      R_o[6,22] := 0.43332982;
      R_o[6,23] := -0.19467659;
      R_o[6,24] := 0.93978935;
      R_o[6,25] := -0.61547863;
      R_o[6,26] := 0.14545523;
      R_o[6,27] := -0.42827970;
      R_o[6,28] := 0.01864699;
      R_o[6,29] := 0.37515923;
      R_o[6,30] := 0.31723750;
      R_o[6,31] := 0.19122434;
      R_o[7,0] := 0.34065035;
      R_o[7,1] := 0.47401485;
      R_o[7,2] := -0.54076427;
      R_o[7,3] := -0.65568548;
      R_o[7,4] := 0.62105906;
      R_o[7,5] := -0.41220605;
      R_o[7,6] := -1.31112802;
      R_o[7,7] := 1.04505157;
      R_o[7,8] := 0.78872794;
      R_o[7,9] := -0.66649288;
      R_o[7,10] := 0.23619340;
      R_o[7,11] := -0.44383812;
      R_o[7,12] := -0.33296376;
      R_o[7,13] := -0.63825399;
      R_o[7,14] := 0.15134087;
      R_o[7,15] := 0.07716195;
      R_o[7,16] := 0.30484754;
      R_o[7,17] := -0.49967739;
      R_o[7,18] := -0.55375117;
      R_o[7,19] := -0.01412584;
      R_o[7,20] := -0.09337062;
      R_o[7,21] := -0.86438709;
      R_o[7,22] := 1.12174129;
      R_o[7,23] := -0.52289206;
      R_o[7,24] := 2.45863652;
      R_o[7,25] := -0.49099314;
      R_o[7,26] := 0.05714682;
      R_o[7,27] := -0.59038329;
      R_o[7,28] := -0.21783109;
      R_o[7,29] := 0.31133965;
      R_o[7,30] := 0.41102508;
      R_o[7,31] := 0.54280049;
      R_o[8,0] := 0.20045589;
      R_o[8,1] := 0.50244647;
      R_o[8,2] := -0.51556474;
      R_o[8,3] := -0.81008476;
      R_o[8,4] := 0.92952043;
      R_o[8,5] := -0.15610516;
      R_o[8,6] := -0.14775947;
      R_o[8,7] := -0.40649518;
      R_o[8,8] := 1.07194042;
      R_o[8,9] := -0.58189887;
      R_o[8,10] := 0.34218273;
      R_o[8,11] := -0.43635336;
      R_o[8,12] := -0.19688728;
      R_o[8,13] := -0.17332749;
      R_o[8,14] := 0.13037777;
      R_o[8,15] := 0.53576058;
      R_o[8,16] := -0.20822550;
      R_o[8,17] := -0.87431055;
      R_o[8,18] := -0.43827292;
      R_o[8,19] := 0.10151042;
      R_o[8,20] := -0.02924687;
      R_o[8,21] := -0.77477866;
      R_o[8,22] := 0.19584732;
      R_o[8,23] := -0.08636574;
      R_o[8,24] := 0.41095579;
      R_o[8,25] := -0.18019967;
      R_o[8,26] := 0.16473477;
      R_o[8,27] := -0.17792331;
      R_o[8,28] := -0.08596105;
      R_o[8,29] := 0.59257406;
      R_o[8,30] := 0.50818813;
      R_o[8,31] := -0.01205147;
      R_o[9,0] := 0.09369560;
      R_o[9,1] := -0.16206230;
      R_o[9,2] := -1.01217055;
      R_o[9,3] := -0.49272183;
      R_o[9,4] := 0.42273074;
      R_o[9,5] := -1.25912929;
      R_o[9,6] := -1.23285043;
      R_o[9,7] := -0.67148495;
      R_o[9,8] := 2.05958033;
      R_o[9,9] := 0.90271044;
      R_o[9,10] := 0.62281978;
      R_o[9,11] := 0.02608189;
      R_o[9,12] := 0.37196815;
      R_o[9,13] := -0.09634275;
      R_o[9,14] := 0.00955611;
      R_o[9,15] := 0.45335814;
      R_o[9,16] := -0.03960776;
      R_o[9,17] := -0.32377270;
      R_o[9,18] := -0.20143498;
      R_o[9,19] := -0.11493812;
      R_o[9,20] := 0.16121885;
      R_o[9,21] := -0.83840460;
      R_o[9,22] := 2.03339243;
      R_o[9,23] := 0.01112972;
      R_o[9,24] := 0.97674733;
      R_o[9,25] := -0.07987648;
      R_o[9,26] := -0.01916505;
      R_o[9,27] := 0.04041042;
      R_o[9,28] := -0.68464011;
      R_o[9,29] := 0.79779410;
      R_o[9,30] := 0.05652495;
      R_o[9,31] := 1.71702218;
      R_o[10,0] := 0.02779424;
      R_o[10,1] := -0.40141207;
      R_o[10,2] := -0.68689167;
      R_o[10,3] := -0.02245888;
      R_o[10,4] := -0.37881848;
      R_o[10,5] := -0.43561807;
      R_o[10,6] := -0.26771024;
      R_o[10,7] := 0.00021951;
      R_o[10,8] := 0.04696209;
      R_o[10,9] := -0.68788171;
      R_o[10,10] := -1.13438833;
      R_o[10,11] := 0.01086713;
      R_o[10,12] := -0.53196830;
      R_o[10,13] := 0.19594459;
      R_o[10,14] := 0.25793335;
      R_o[10,15] := -0.32604316;
      R_o[10,16] := 0.37373966;
      R_o[10,17] := -0.17519239;
      R_o[10,18] := -0.50413275;
      R_o[10,19] := -0.21772946;
      R_o[10,20] := -0.45339233;
      R_o[10,21] := -0.80154604;
      R_o[10,22] := 1.25618088;
      R_o[10,23] := -0.80704057;
      R_o[10,24] := 0.59909791;
      R_o[10,25] := 0.20229515;
      R_o[10,26] := 0.21944004;
      R_o[10,27] := -0.56646466;
      R_o[10,28] := -0.31041694;
      R_o[10,29] := 0.22589801;
      R_o[10,30] := -0.05355195;
      R_o[10,31] := 0.32136935;
      R_o[11,0] := 0.13318552;
      R_o[11,1] := 0.14860928;
      R_o[11,2] := -1.01276350;
      R_o[11,3] := -0.72060043;
      R_o[11,4] := 0.21185312;
      R_o[11,5] := -0.54846334;
      R_o[11,6] := -0.80948603;
      R_o[11,7] := -0.51698428;
      R_o[11,8] := 0.54447424;
      R_o[11,9] := -0.08923292;
      R_o[11,10] := 0.80089408;
      R_o[11,11] := -0.46713293;
      R_o[11,12] := -0.18385221;
      R_o[11,13] := -0.25236073;
      R_o[11,14] := -0.38691062;
      R_o[11,15] := 0.41189039;
      R_o[11,16] := -0.15554635;
      R_o[11,17] := -0.20958538;
      R_o[11,18] := -0.33747688;
      R_o[11,19] := -0.01130310;
      R_o[11,20] := -0.34684128;
      R_o[11,21] := -1.16357529;
      R_o[11,22] := 0.93542528;
      R_o[11,23] := -0.32925424;
      R_o[11,24] := -0.24023592;
      R_o[11,25] := 0.18446164;
      R_o[11,26] := 0.29880688;
      R_o[11,27] := -0.74903917;
      R_o[11,28] := -0.72029477;
      R_o[11,29] := 0.05337867;
      R_o[11,30] := 0.33378384;
      R_o[11,31] := 0.49327818;
      R_o[12,0] := -0.20777129;
      R_o[12,1] := 0.40653828;
      R_o[12,2] := -1.15580094;
      R_o[12,3] := -0.58007532;
      R_o[12,4] := 0.60843307;
      R_o[12,5] := -0.29073319;
      R_o[12,6] := -1.30077088;
      R_o[12,7] := -0.48383486;
      R_o[12,8] := 0.50866872;
      R_o[12,9] := -0.32799762;
      R_o[12,10] := 0.08853685;
      R_o[12,11] := -0.12722090;
      R_o[12,12] := -0.13251597;
      R_o[12,13] := -0.53875893;
      R_o[12,14] := 0.53165895;
      R_o[12,15] := -0.15170568;
      R_o[12,16] := 0.36354136;
      R_o[12,17] := -0.40015194;
      R_o[12,18] := -0.16225255;
      R_o[12,19] := 0.10627833;
      R_o[12,20] := -0.51227063;
      R_o[12,21] := -1.87520730;
      R_o[12,22] := 0.45057613;
      R_o[12,23] := -0.53412980;
      R_o[12,24] := 1.92583394;
      R_o[12,25] := -0.02440960;
      R_o[12,26] := -0.29421479;
      R_o[12,27] := -0.31305516;
      R_o[12,28] := -0.33143687;
      R_o[12,29] := 0.62461257;
      R_o[12,30] := -0.20750031;
      R_o[12,31] := -0.49445149;
      R_o[13,0] := 0.03614095;
      R_o[13,1] := 0.71849424;
      R_o[13,2] := -0.54970086;
      R_o[13,3] := -1.13958406;
      R_o[13,4] := 0.13165674;
      R_o[13,5] := -0.29205301;
      R_o[13,6] := -0.17687124;
      R_o[13,7] := -0.44388226;
      R_o[13,8] := 0.55644709;
      R_o[13,9] := -1.64114189;
      R_o[13,10] := 0.36598471;
      R_o[13,11] := -0.55834091;
      R_o[13,12] := -0.65976113;
      R_o[13,13] := -0.56921744;
      R_o[13,14] := 0.36256570;
      R_o[13,15] := 0.93002528;
      R_o[13,16] := 0.01155506;
      R_o[13,17] := -1.06603146;
      R_o[13,18] := -0.26420283;
      R_o[13,19] := 0.73663074;
      R_o[13,20] := 0.70005757;
      R_o[13,21] := -2.01711774;
      R_o[13,22] := 1.58053350;
      R_o[13,23] := -0.36436135;
      R_o[13,24] := 1.53379405;
      R_o[13,25] := -0.02658881;
      R_o[13,26] := -0.55448914;
      R_o[13,27] := -0.54852170;
      R_o[13,28] := -0.88863921;
      R_o[13,29] := 0.60738230;
      R_o[13,30] := 0.84559155;
      R_o[13,31] := 0.56188303;
      R_o[14,0] := 0.01524067;
      R_o[14,1] := -0.33807415;
      R_o[14,2] := -0.05662629;
      R_o[14,3] := -0.35284707;
      R_o[14,4] := -0.61716205;
      R_o[14,5] := 0.14316405;
      R_o[14,6] := -0.07415292;
      R_o[14,7] := 0.05172193;
      R_o[14,8] := -0.41683775;
      R_o[14,9] := 0.26181215;
      R_o[14,10] := -0.04171603;
      R_o[14,11] := -0.11402290;
      R_o[14,12] := 0.21671122;
      R_o[14,13] := -0.58848882;
      R_o[14,14] := -1.07252192;
      R_o[14,15] := -0.00347600;
      R_o[14,16] := -0.06543477;
      R_o[14,17] := 0.08887091;
      R_o[14,18] := -0.26554459;
      R_o[14,19] := 0.10296860;
      R_o[14,20] := -0.15775499;
      R_o[14,21] := -0.13629206;
      R_o[14,22] := 0.34778851;
      R_o[14,23] := 0.24370442;
      R_o[14,24] := 0.21042643;
      R_o[14,25] := -0.39436981;
      R_o[14,26] := 0.31873849;
      R_o[14,27] := -0.23981427;
      R_o[14,28] := -0.30328980;
      R_o[14,29] := 0.43482566;
      R_o[14,30] := 0.04193076;
      R_o[14,31] := -0.31264323;
      R_o[15,0] := 0.29360059;
      R_o[15,1] := 0.36706486;
      R_o[15,2] := -0.51066637;
      R_o[15,3] := -0.09302752;
      R_o[15,4] := 0.32202122;
      R_o[15,5] := -0.14361922;
      R_o[15,6] := -0.80344599;
      R_o[15,7] := 0.33518144;
      R_o[15,8] := -0.17809442;
      R_o[15,9] := -0.02201664;
      R_o[15,10] := 0.29279521;
      R_o[15,11] := -0.10687640;
      R_o[15,12] := -0.69306546;
      R_o[15,13] := -0.34347835;
      R_o[15,14] := 0.21410543;
      R_o[15,15] := -1.83093214;
      R_o[15,16] := -0.11691079;
      R_o[15,17] := -0.45732704;
      R_o[15,18] := -0.86807251;
      R_o[15,19] := 0.23608641;
      R_o[15,20] := 0.10597400;
      R_o[15,21] := 0.15834263;
      R_o[15,22] := 0.78955311;
      R_o[15,23] := -0.16079797;
      R_o[15,24] := 0.00513626;
      R_o[15,25] := -0.28376704;
      R_o[15,26] := 0.66462660;
      R_o[15,27] := -0.28953049;
      R_o[15,28] := 0.16934998;
      R_o[15,29] := -0.14268929;
      R_o[15,30] := -0.18818894;
      R_o[15,31] := 0.12157705;
      R_o[16,0] := 0.07833512;
      R_o[16,1] := 0.23961815;
      R_o[16,2] := -0.40951693;
      R_o[16,3] := -0.29096887;
      R_o[16,4] := 0.11224928;
      R_o[16,5] := -0.50798362;
      R_o[16,6] := -0.34913379;
      R_o[16,7] := 0.10367194;
      R_o[16,8] := 0.61167037;
      R_o[16,9] := -0.11267250;
      R_o[16,10] := 0.56287217;
      R_o[16,11] := -0.03040320;
      R_o[16,12] := 0.23440740;
      R_o[16,13] := -0.01905249;
      R_o[16,14] := -0.25718442;
      R_o[16,15] := 0.23948520;
      R_o[16,16] := -0.43410707;
      R_o[16,17] := -0.35836715;
      R_o[16,18] := 0.24731942;
      R_o[16,19] := -0.06834326;
      R_o[16,20] := -0.08543305;
      R_o[16,21] := -0.02655645;
      R_o[16,22] := 0.59191698;
      R_o[16,23] := -0.21830332;
      R_o[16,24] := -0.06442533;
      R_o[16,25] := 0.02223889;
      R_o[16,26] := 0.14285798;
      R_o[16,27] := 0.25474730;
      R_o[16,28] := -0.40410686;
      R_o[16,29] := 0.24501032;
      R_o[16,30] := -0.03571527;
      R_o[16,31] := -0.42208397;
      R_o[17,0] := 0.15439741;
      R_o[17,1] := -0.02684163;
      R_o[17,2] := -0.32831976;
      R_o[17,3] := -0.36610043;
      R_o[17,4] := 0.24014680;
      R_o[17,5] := 0.02118563;
      R_o[17,6] := 0.24636027;
      R_o[17,7] := -0.17018878;
      R_o[17,8] := 0.02465408;
      R_o[17,9] := 0.45513898;
      R_o[17,10] := 0.80733585;
      R_o[17,11] := 0.14326459;
      R_o[17,12] := 0.49080721;
      R_o[17,13] := -0.27932650;
      R_o[17,14] := -0.49028867;
      R_o[17,15] := 0.32682586;
      R_o[17,16] := -0.48414201;
      R_o[17,17] := 0.85723203;
      R_o[17,18] := 0.24715909;
      R_o[17,19] := 0.22189638;
      R_o[17,20] := -0.06566357;
      R_o[17,21] := 0.11126448;
      R_o[17,22] := 0.06685662;
      R_o[17,23] := 0.21587326;
      R_o[17,24] := 0.30921510;
      R_o[17,25] := 0.01129790;
      R_o[17,26] := 0.09004966;
      R_o[17,27] := -0.09074225;
      R_o[17,28] := -0.03670594;
      R_o[17,29] := -0.11644791;
      R_o[17,30] := -0.05028833;
      R_o[17,31] := -0.26572007;
      R_o[18,0] := 0.84484732;
      R_o[18,1] := 0.53163010;
      R_o[18,2] := 0.00904752;
      R_o[18,3] := -0.46008062;
      R_o[18,4] := -0.02926146;
      R_o[18,5] := -0.21939951;
      R_o[18,6] := -0.28743288;
      R_o[18,7] := 0.18235296;
      R_o[18,8] := -0.05455190;
      R_o[18,9] := -0.52153742;
      R_o[18,10] := -0.11111192;
      R_o[18,11] := -0.24852699;
      R_o[18,12] := 0.08671411;
      R_o[18,13] := -0.15882707;
      R_o[18,14] := 0.04479800;
      R_o[18,15] := 0.31299874;
      R_o[18,16] := -0.02502846;
      R_o[18,17] := -0.62176991;
      R_o[18,18] := 0.53988975;
      R_o[18,19] := -0.09278865;
      R_o[18,20] := 0.15000486;
      R_o[18,21] := -0.30583379;
      R_o[18,22] := -0.07494947;
      R_o[18,23] := -0.04273816;
      R_o[18,24] := -0.03186971;
      R_o[18,25] := -0.37590668;
      R_o[18,26] := 0.54982477;
      R_o[18,27] := -0.21423021;
      R_o[18,28] := -0.32949436;
      R_o[18,29] := 0.24937831;
      R_o[18,30] := 0.11211216;
      R_o[18,31] := 0.24685173;
      R_o[19,0] := 0.10862272;
      R_o[19,1] := 0.48960793;
      R_o[19,2] := 0.00677478;
      R_o[19,3] := -0.79965466;
      R_o[19,4] := 0.39394405;
      R_o[19,5] := 0.38277546;
      R_o[19,6] := -0.18124942;
      R_o[19,7] := -0.22815390;
      R_o[19,8] := 1.09245586;
      R_o[19,9] := -0.67992783;
      R_o[19,10] := 0.28631067;
      R_o[19,11] := -0.19220580;
      R_o[19,12] := 0.50091755;
      R_o[19,13] := -0.70053983;
      R_o[19,14] := -0.24056637;
      R_o[19,15] := 0.44088650;
      R_o[19,16] := -0.03423277;
      R_o[19,17] := 0.15923414;
      R_o[19,18] := -0.11861752;
      R_o[19,19] := 0.20712623;
      R_o[19,20] := 0.05342558;
      R_o[19,21] := -0.45508027;
      R_o[19,22] := 0.20025966;
      R_o[19,23] := -0.11695480;
      R_o[19,24] := 0.66766268;
      R_o[19,25] := -0.57887745;
      R_o[19,26] := 0.04404074;
      R_o[19,27] := -0.37624091;
      R_o[19,28] := -0.39110780;
      R_o[19,29] := 0.61437207;
      R_o[19,30] := 0.16036567;
      R_o[19,31] := 0.27669203;
      R_o[20,0] := -0.01197398;
      R_o[20,1] := 0.27682754;
      R_o[20,2] := -1.47277486;
      R_o[20,3] := -0.79019433;
      R_o[20,4] := 0.34979358;
      R_o[20,5] := -0.53736645;
      R_o[20,6] := -1.85887754;
      R_o[20,7] := -0.42141077;
      R_o[20,8] := -0.63334978;
      R_o[20,9] := -0.62121934;
      R_o[20,10] := 0.47573924;
      R_o[20,11] := -0.12207225;
      R_o[20,12] := 0.12717439;
      R_o[20,13] := -0.79209167;
      R_o[20,14] := -0.06180368;
      R_o[20,15] := 0.27822039;
      R_o[20,16] := 0.00291310;
      R_o[20,17] := -0.25131065;
      R_o[20,18] := -0.09981156;
      R_o[20,19] := 0.25378519;
      R_o[20,20] := -1.01099992;
      R_o[20,21] := -1.39382052;
      R_o[20,22] := 0.59680003;
      R_o[20,23] := -0.44065499;
      R_o[20,24] := 1.74228501;
      R_o[20,25] := -0.03751455;
      R_o[20,26] := -0.60711169;
      R_o[20,27] := -0.39512217;
      R_o[20,28] := -0.13597757;
      R_o[20,29] := 0.10179781;
      R_o[20,30] := 0.42191899;
      R_o[20,31] := 0.58368075;
      R_o[21,0] := -0.24594249;
      R_o[21,1] := 0.04108999;
      R_o[21,2] := -0.60767484;
      R_o[21,3] := -0.60254490;
      R_o[21,4] := 0.06250022;
      R_o[21,5] := -0.14623532;
      R_o[21,6] := -0.28648895;
      R_o[21,7] := -0.01256131;
      R_o[21,8] := 0.55629826;
      R_o[21,9] := -0.27424589;
      R_o[21,10] := 0.43336782;
      R_o[21,11] := -0.08429422;
      R_o[21,12] := -0.15243714;
      R_o[21,13] := -0.45141295;
      R_o[21,14] := 0.12675479;
      R_o[21,15] := -0.09365185;
      R_o[21,16] := 0.27947018;
      R_o[21,17] := -0.34975228;
      R_o[21,18] := -0.28150943;
      R_o[21,19] := -0.03043183;
      R_o[21,20] := -0.22126247;
      R_o[21,21] := -0.01680325;
      R_o[21,22] := 0.48534319;
      R_o[21,23] := -0.07723329;
      R_o[21,24] := 0.63475794;
      R_o[21,25] := 0.04629425;
      R_o[21,26] := 0.04529271;
      R_o[21,27] := -0.37165093;
      R_o[21,28] := -0.13515891;
      R_o[21,29] := 0.46588650;
      R_o[21,30] := 0.48834196;
      R_o[21,31] := 0.07594018;
      R_o[22,0] := 0.27011484;
      R_o[22,1] := 0.40486771;
      R_o[22,2] := -0.28902775;
      R_o[22,3] := -0.48784915;
      R_o[22,4] := 0.28023198;
      R_o[22,5] := -0.34532472;
      R_o[22,6] := -0.53983426;
      R_o[22,7] := -0.54445738;
      R_o[22,8] := 0.08511036;
      R_o[22,9] := -0.25733194;
      R_o[22,10] := 0.29259899;
      R_o[22,11] := -0.16682011;
      R_o[22,12] := -0.45611075;
      R_o[22,13] := -0.06053562;
      R_o[22,14] := -0.93061149;
      R_o[22,15] := -0.12850389;
      R_o[22,16] := -0.21759163;
      R_o[22,17] := -0.33520815;
      R_o[22,18] := -0.21541405;
      R_o[22,19] := 0.05377239;
      R_o[22,20] := -0.23695599;
      R_o[22,21] := 0.01863871;
      R_o[22,22] := 0.46674144;
      R_o[22,23] := -0.05650645;
      R_o[22,24] := 0.71159017;
      R_o[22,25] := -0.32194561;
      R_o[22,26] := -0.34680220;
      R_o[22,27] := -0.28244287;
      R_o[22,28] := 0.15536174;
      R_o[22,29] := -0.16343887;
      R_o[22,30] := 0.10497386;
      R_o[22,31] := 0.53858823;
      R_o[23,0] := 0.34600383;
      R_o[23,1] := 0.42481279;
      R_o[23,2] := 0.07165840;
      R_o[23,3] := -0.50042599;
      R_o[23,4] := 0.28742552;
      R_o[23,5] := 0.16970187;
      R_o[23,6] := 0.16972134;
      R_o[23,7] := 0.16999744;
      R_o[23,8] := 0.32839668;
      R_o[23,9] := -0.02685527;
      R_o[23,10] := -0.00342671;
      R_o[23,11] := -0.28909808;
      R_o[23,12] := 0.03453528;
      R_o[23,13] := -0.30969155;
      R_o[23,14] := 0.31023362;
      R_o[23,15] := 0.13957487;
      R_o[23,16] := 0.17285080;
      R_o[23,17] := -0.09276348;
      R_o[23,18] := -0.32455254;
      R_o[23,19] := 0.16625991;
      R_o[23,20] := -0.04450256;
      R_o[23,21] := -0.23909336;
      R_o[23,22] := 0.36995435;
      R_o[23,23] := -0.37734264;
      R_o[23,24] := 0.42270988;
      R_o[23,25] := -0.30175060;
      R_o[23,26] := 0.09778602;
      R_o[23,27] := -0.68427491;
      R_o[23,28] := -0.12598298;
      R_o[23,29] := 0.25889975;
      R_o[23,30] := 0.37449488;
      R_o[23,31] := 0.03907451;
      R_o[24,0] := 0.20198651;
      R_o[24,1] := 0.36463314;
      R_o[24,2] := -0.31008822;
      R_o[24,3] := -0.05163987;
      R_o[24,4] := 0.28869891;
      R_o[24,5] := 0.01050948;
      R_o[24,6] := -0.20344213;
      R_o[24,7] := -0.25559375;
      R_o[24,8] := 0.31342509;
      R_o[24,9] := -0.41931885;
      R_o[24,10] := -0.02418928;
      R_o[24,11] := -0.32550445;
      R_o[24,12] := -0.49690139;
      R_o[24,13] := -0.44138038;
      R_o[24,14] := -0.04818862;
      R_o[24,15] := 0.49021626;
      R_o[24,16] := 0.01580368;
      R_o[24,17] := -0.74874520;
      R_o[24,18] := -0.06684852;
      R_o[24,19] := 0.50041729;
      R_o[24,20] := -0.22713709;
      R_o[24,21] := -0.22028215;
      R_o[24,22] := 0.25357047;
      R_o[24,23] := -0.44678640;
      R_o[24,24] := -0.33140028;
      R_o[24,25] := -0.19499658;
      R_o[24,26] := 0.01837249;
      R_o[24,27] := -0.17397606;
      R_o[24,28] := -0.37122267;
      R_o[24,29] := 0.10083988;
      R_o[24,30] := 0.41414759;
      R_o[24,31] := 0.16101778;
      R_o[25,0] := 0.05109156;
      R_o[25,1] := 0.13809530;
      R_o[25,2] := -0.42768860;
      R_o[25,3] := -0.46329850;
      R_o[25,4] := -0.01765707;
      R_o[25,5] := -0.01810573;
      R_o[25,6] := -0.22468179;
      R_o[25,7] := 0.17521209;
      R_o[25,8] := 0.34461039;
      R_o[25,9] := -0.11726221;
      R_o[25,10] := 0.49146181;
      R_o[25,11] := 0.27963191;
      R_o[25,12] := 0.37571144;
      R_o[25,13] := -0.02800122;
      R_o[25,14] := -0.22924468;
      R_o[25,15] := -0.03784134;
      R_o[25,16] := -0.12258809;
      R_o[25,17] := -0.31369281;
      R_o[25,18] := -0.21762075;
      R_o[25,19] := -0.23435897;
      R_o[25,20] := -0.26502833;
      R_o[25,21] := 0.18020962;
      R_o[25,22] := 0.09507836;
      R_o[25,23] := -0.08545585;
      R_o[25,24] := 0.48384097;
      R_o[25,25] := 0.22817534;
      R_o[25,26] := -0.26306638;
      R_o[25,27] := -0.15757905;
      R_o[25,28] := -0.20556410;
      R_o[25,29] := 0.62218368;
      R_o[25,30] := 0.10382322;
      R_o[25,31] := 0.02228775;
      R_o[26,0] := 0.04785801;
      R_o[26,1] := 0.15561581;
      R_o[26,2] := 0.22885913;
      R_o[26,3] := -0.60473061;
      R_o[26,4] := 0.47135803;
      R_o[26,5] := -0.33018327;
      R_o[26,6] := -1.03677499;
      R_o[26,7] := -0.22189558;
      R_o[26,8] := -0.13217314;
      R_o[26,9] := -0.01338464;
      R_o[26,10] := 0.64015561;
      R_o[26,11] := -0.13306759;
      R_o[26,12] := 0.19538191;
      R_o[26,13] := -1.67280841;
      R_o[26,14] := -0.12914124;
      R_o[26,15] := 0.51318997;
      R_o[26,16] := 0.29180083;
      R_o[26,17] := -0.37431264;
      R_o[26,18] := -0.20381257;
      R_o[26,19] := 0.61842877;
      R_o[26,20] := -0.43941274;
      R_o[26,21] := -3.21122694;
      R_o[26,22] := 2.21060944;
      R_o[26,23] := -0.29611194;
      R_o[26,24] := 4.76488018;
      R_o[26,25] := -0.00677092;
      R_o[26,26] := 0.95254189;
      R_o[26,27] := -0.80067807;
      R_o[26,28] := -0.16087081;
      R_o[26,29] := 0.26623115;
      R_o[26,30] := 0.82952696;
      R_o[26,31] := -1.02879465;
      R_o[27,0] := 0.14549352;
      R_o[27,1] := 0.27596897;
      R_o[27,2] := -0.44747168;
      R_o[27,3] := -0.83414388;
      R_o[27,4] := 0.31795341;
      R_o[27,5] := -0.90306568;
      R_o[27,6] := -0.42387462;
      R_o[27,7] := 0.02974604;
      R_o[27,8] := 1.84534919;
      R_o[27,9] := -0.65307516;
      R_o[27,10] := 0.66818446;
      R_o[27,11] := -0.02700442;
      R_o[27,12] := -0.91477334;
      R_o[27,13] := -0.66135025;
      R_o[27,14] := -0.10455511;
      R_o[27,15] := 0.00713633;
      R_o[27,16] := -0.19336109;
      R_o[27,17] := -0.34954131;
      R_o[27,18] := -0.23724046;
      R_o[27,19] := -0.44211617;
      R_o[27,20] := -0.00597036;
      R_o[27,21] := -1.56280470;
      R_o[27,22] := 0.64400321;
      R_o[27,23] := -0.45753676;
      R_o[27,24] := -0.28298530;
      R_o[27,25] := 0.30139643;
      R_o[27,26] := 0.44311312;
      R_o[27,27] := -1.28934312;
      R_o[27,28] := -0.27950504;
      R_o[27,29] := -0.03651794;
      R_o[27,30] := 0.23414747;
      R_o[27,31] := 0.66848058;
      R_o[28,0] := 0.10052842;
      R_o[28,1] := 0.95776904;
      R_o[28,2] := -0.58687061;
      R_o[28,3] := -0.52412993;
      R_o[28,4] := 0.28911093;
      R_o[28,5] := -0.93690294;
      R_o[28,6] := -0.44405863;
      R_o[28,7] := -0.39684597;
      R_o[28,8] := 0.22224870;
      R_o[28,9] := -0.50384551;
      R_o[28,10] := 0.44301915;
      R_o[28,11] := -0.25398868;
      R_o[28,12] := -0.45412725;
      R_o[28,13] := 0.03549762;
      R_o[28,14] := -0.04904316;
      R_o[28,15] := 0.08361682;
      R_o[28,16] := -0.12424450;
      R_o[28,17] := -0.14209995;
      R_o[28,18] := -0.02077562;
      R_o[28,19] := 0.33017302;
      R_o[28,20] := -0.21900289;
      R_o[28,21] := -0.28608552;
      R_o[28,22] := 1.11653757;
      R_o[28,23] := -0.20174463;
      R_o[28,24] := 1.74418199;
      R_o[28,25] := -0.11653454;
      R_o[28,26] := 0.26567152;
      R_o[28,27] := 0.18579985;
      R_o[28,28] := 0.05587514;
      R_o[28,29] := 1.14281774;
      R_o[28,30] := 0.14929593;
      R_o[28,31] := 0.15964474;
      R_o[29,0] := 0.07655234;
      R_o[29,1] := 0.00526063;
      R_o[29,2] := -0.60426944;
      R_o[29,3] := -0.67821729;
      R_o[29,4] := 0.48224354;
      R_o[29,5] := 0.24618737;
      R_o[29,6] := -1.01446080;
      R_o[29,7] := -0.21527001;
      R_o[29,8] := 0.31270966;
      R_o[29,9] := -0.64469713;
      R_o[29,10] := 0.30272844;
      R_o[29,11] := -0.49371287;
      R_o[29,12] := -0.25839141;
      R_o[29,13] := -0.60940570;
      R_o[29,14] := 0.23404275;
      R_o[29,15] := 0.34532225;
      R_o[29,16] := 0.00867103;
      R_o[29,17] := -0.31875700;
      R_o[29,18] := -0.37785101;
      R_o[29,19] := -0.11795938;
      R_o[29,20] := -0.80922771;
      R_o[29,21] := -0.48978224;
      R_o[29,22] := 1.59050429;
      R_o[29,23] := -0.40486097;
      R_o[29,24] := 1.31220138;
      R_o[29,25] := -0.15769550;
      R_o[29,26] := -0.18835722;
      R_o[29,27] := -0.71010518;
      R_o[29,28] := 0.08438613;
      R_o[29,29] := -0.27337590;
      R_o[29,30] := 0.64987278;
      R_o[29,31] := -0.28353274;
      R_o[30,0] := -0.04396043;
      R_o[30,1] := -0.50152326;
      R_o[30,2] := -0.45781407;
      R_o[30,3] := -0.94959831;
      R_o[30,4] := 0.37568477;
      R_o[30,5] := -3.20458865;
      R_o[30,6] := -0.45303726;
      R_o[30,7] := -0.21864329;
      R_o[30,8] := 3.02453923;
      R_o[30,9] := -1.07397604;
      R_o[30,10] := 0.58351398;
      R_o[30,11] := -0.24423414;
      R_o[30,12] := -0.56096327;
      R_o[30,13] := -0.16615988;
      R_o[30,14] := -0.17139067;
      R_o[30,15] := 0.10854375;
      R_o[30,16] := -0.12342630;
      R_o[30,17] := -0.58460224;
      R_o[30,18] := -0.26377097;
      R_o[30,19] := 1.32042170;
      R_o[30,20] := -0.53046167;
      R_o[30,21] := -3.48458099;
      R_o[30,22] := 1.21924889;
      R_o[30,23] := -0.29753938;
      R_o[30,24] := 0.52615410;
      R_o[30,25] := -0.07486701;
      R_o[30,26] := 0.17118107;
      R_o[30,27] := -0.52948815;
      R_o[30,28] := -0.66240865;
      R_o[30,29] := 0.88388693;
      R_o[30,30] := 1.60189033;
      R_o[30,31] := -0.25331134;
      R_o[31,0] := -0.29912165;
      R_o[31,1] := 0.42477793;
      R_o[31,2] := -0.21023647;
      R_o[31,3] := -0.11975008;
      R_o[31,4] := -0.01268277;
      R_o[31,5] := -0.02130502;
      R_o[31,6] := 0.03439108;
      R_o[31,7] := 0.05758012;
      R_o[31,8] := 0.41448206;
      R_o[31,9] := -0.14623728;
      R_o[31,10] := -0.23915647;
      R_o[31,11] := 0.37064037;
      R_o[31,12] := 0.17834072;
      R_o[31,13] := -0.36577532;
      R_o[31,14] := 0.50369042;
      R_o[31,15] := 0.49751189;
      R_o[31,16] := 0.05057595;
      R_o[31,17] := -0.61116600;
      R_o[31,18] := -0.19325699;
      R_o[31,19] := -0.20192310;
      R_o[31,20] := -0.16053063;
      R_o[31,21] := -0.19299865;
      R_o[31,22] := 0.76509267;
      R_o[31,23] := -0.20398943;
      R_o[31,24] := 0.69476819;
      R_o[31,25] := -0.17712449;
      R_o[31,26] := -0.27581781;
      R_o[31,27] := -0.35418263;
      R_o[31,28] := -0.04145564;
      R_o[31,29] := 0.11614407;
      R_o[31,30] := 0.36519545;
      R_o[31,31] := 0.51034522;
      B_i[0] := 0.29052719;
      B_i[1] := 0.13999742;
      B_i[2] := 0.05400676;
      B_i[3] := 1.21956277;
      B_i[4] := 0.53838974;
      B_i[5] := 0.34135109;
      B_i[6] := 0.58119547;
      B_i[7] := 0.72373772;
      B_i[8] := 0.18965542;
      B_i[9] := 0.22784001;
      B_i[10] := 0.12681076;
      B_i[11] := -0.31453860;
      B_i[12] := 0.99506211;
      B_i[13] := -0.25184420;
      B_i[14] := 0.57154953;
      B_i[15] := 0.68310666;
      B_i[16] := 0.46907067;
      B_i[17] := 1.38582957;
      B_i[18] := 0.21330455;
      B_i[19] := 0.55320585;
      B_i[20] := 0.14247677;
      B_i[21] := 1.30028939;
      B_i[22] := -0.03355794;
      B_i[23] := 0.97606659;
      B_i[24] := -0.32917467;
      B_i[25] := 0.11296137;
      B_i[26] := 0.60575831;
      B_i[27] := 0.12289220;
      B_i[28] := 0.12378435;
      B_i[29] := -0.20421156;
      B_i[30] := 2.04777122;
      B_i[31] := 0.58692878;
      B_f[0] := 0.59489554;
      B_f[1] := 1.40699565;
      B_f[2] := 2.19698429;
      B_f[3] := -2.09258509;
      B_f[4] := -0.35761544;
      B_f[5] := 1.81703711;
      B_f[6] := -0.20773043;
      B_f[7] := 0.08518680;
      B_f[8] := 1.02957809;
      B_f[9] := 0.39947632;
      B_f[10] := -0.41881144;
      B_f[11] := -0.18117729;
      B_f[12] := 0.60140902;
      B_f[13] := 2.14849520;
      B_f[14] := -0.99196982;
      B_f[15] := 0.14013851;
      B_f[16] := -0.17579740;
      B_f[17] := -0.68764311;
      B_f[18] := 0.13257200;
      B_f[19] := 1.12185311;
      B_f[20] := 2.08465552;
      B_f[21] := -1.33065128;
      B_f[22] := 1.84940779;
      B_f[23] := -0.39349115;
      B_f[24] := 1.96590114;
      B_f[25] := -0.18333542;
      B_f[26] := 1.47585058;
      B_f[27] := -0.81844461;
      B_f[28] := 1.81535029;
      B_f[29] := -0.78683877;
      B_f[30] := 0.60889250;
      B_f[31] := 0.83791882;
      B_g[0] := 0.22905608;
      B_g[1] := 0.17009147;
      B_g[2] := -0.48756313;
      B_g[3] := -1.28816998;
      B_g[4] := 0.67155010;
      B_g[5] := -0.28815305;
      B_g[6] := -0.53673601;
      B_g[7] := 0.18329665;
      B_g[8] := 0.26111066;
      B_g[9] := -0.47462666;
      B_g[10] := 0.24001265;
      B_g[11] := 0.08113776;
      B_g[12] := 0.26064369;
      B_g[13] := -0.50959384;
      B_g[14] := 0.13000551;
      B_g[15] := 0.03399255;
      B_g[16] := -0.05519996;
      B_g[17] := -1.02396870;
      B_g[18] := -0.65365821;
      B_g[19] := 0.52074474;
      B_g[20] := 0.07321863;
      B_g[21] := -0.85776556;
      B_g[22] := 0.20937879;
      B_g[23] := -0.20943075;
      B_g[24] := 0.58523530;
      B_g[25] := -0.22898147;
      B_g[26] := -0.04568266;
      B_g[27] := -0.53164268;
      B_g[28] := -0.86436212;
      B_g[29] := 0.15611494;
      B_g[30] := 0.35011026;
      B_g[31] := 0.19370955;
      B_o[0] := 1.49208975;
      B_o[1] := 2.81516886;
      B_o[2] := 2.18883061;
      B_o[3] := -0.09973972;
      B_o[4] := 1.51783991;
      B_o[5] := 2.80428600;
      B_o[6] := 1.25245881;
      B_o[7] := 2.54309654;
      B_o[8] := 2.19469237;
      B_o[9] := 3.42261577;
      B_o[10] := 0.69256198;
      B_o[11] := 1.89961219;
      B_o[12] := 2.60195112;
      B_o[13] := 2.74219322;
      B_o[14] := 1.12739038;
      B_o[15] := 0.73841697;
      B_o[16] := 2.09512138;
      B_o[17] := 0.25980064;
      B_o[18] := 1.51229715;
      B_o[19] := 2.18297529;
      B_o[20] := 2.48969460;
      B_o[21] := 2.40099096;
      B_o[22] := 2.13614511;
      B_o[23] := 1.86597776;
      B_o[24] := 1.81434488;
      B_o[25] := 1.40169716;
      B_o[26] := 2.14857674;
      B_o[27] := 1.86558235;
      B_o[28] := 2.20261288;
      B_o[29] := 1.91678286;
      B_o[30] := 2.64595127;
      B_o[31] := 1.97294784;
      FC_W[0,0] := -0.50072664;
      FC_W[0,1] := 0.38558379;
      FC_W[0,2] := -0.35383445;
      FC_W[0,3] := 0.17127538;
      FC_W[0,4] := -0.39166355;
      FC_W[0,5] := 0.57908976;
      FC_W[0,6] := -1.36387634;
      FC_W[0,7] := 1.36579943;
      FC_W[0,8] := -0.32925993;
      FC_W[0,9] := 1.01634562;
      FC_W[0,10] := 0.00445139;
      FC_W[0,11] := 0.69473535;
      FC_W[0,12] := -0.49821049;
      FC_W[0,13] := -0.26812953;
      FC_W[0,14] := 0.26458338;
      FC_W[0,15] := -0.07245288;
      FC_W[0,16] := -0.28500775;
      FC_W[0,17] := -0.39852720;
      FC_W[0,18] := -0.81462759;
      FC_W[0,19] := -0.50401014;
      FC_W[0,20] := 0.98045069;
      FC_W[0,21] := -0.53436071;
      FC_W[0,22] := 1.18371463;
      FC_W[0,23] := 1.13741755;
      FC_W[0,24] := -0.49609959;
      FC_W[0,25] := 0.17210497;
      FC_W[0,26] := -0.13020390;
      FC_W[0,27] := 0.78402209;
      FC_W[0,28] := -0.33053657;
      FC_W[0,29] := 0.29995582;
      FC_W[0,30] := -0.17268366;
      FC_W[0,31] := 0.03926789;
      FC_W[1,0] := 1.05041742;
      FC_W[1,1] := -0.16195486;
      FC_W[1,2] := 0.19831444;
      FC_W[1,3] := 0.04361769;
      FC_W[1,4] := 1.01592088;
      FC_W[1,5] := 1.06561565;
      FC_W[1,6] := 0.50277889;
      FC_W[1,7] := 0.90347242;
      FC_W[1,8] := 0.68030423;
      FC_W[1,9] := -0.20029935;
      FC_W[1,10] := 0.17466098;
      FC_W[1,11] := 0.27924612;
